// Device/Application/ST/ST_MACHINE/ST_MACHINE_PUBLIC
TYPE ST_MACHINE_PUBLIC :
STRUCT
	xEnabled             : BOOL; // Станок включен в работу
	xDisablePending      : BOOL; // Запрошено отключение после выхода автомата в разрешённый шаг
	xPowerAllowed        : BOOL; // Кнопка включения, отключения или отмены отключения доступна
	xResetAllowed        : BOOL; // Кнопка сброса ошибки станка доступна
	xManualControlAllowed       : BOOL; // Ручное управление разрешено режимом и состоянием станка
	xManualSafetyDoorControlEnabled : BOOL; // Операторская дверь управляется только моделью
	xManualSafetyDoorOpenAllowed : BOOL; // Разрешено открыть операторскую дверь
	xManualSafetyDoorCloseAllowed: BOOL; // Разрешено закрыть операторскую дверь
	xManualHatchOpenAllowed      : BOOL; // Разрешено открыть роботный люк
	xManualHatchCloseAllowed     : BOOL; // Разрешено закрыть роботный люк
	xManualHatchUnlockAllowed    : BOOL; // Разрешено открыть замок роботного люка
	xManualHatchLockAllowed      : BOOL; // Разрешено закрыть замок роботного люка
	xManualChuckOpenAllowed      : BOOL; // Разрешено разжать патрон
	xManualChuckCloseAllowed     : BOOL; // Разрешено зажать патрон
	xProcessing          : BOOL; // Станок выполняет цикл обработки
    xPartReady           : BOOL; // Обработка детали завершена
    xServiceRequired     : BOOL; // Станку требуется обслуживание роботом
    xCanAcceptService    : BOOL; // Станок готов принять робота
    xRobotReleased       : BOOL; // Робот освобождён после операции
	xDone                : BOOL; // Операция обслуживания завершена
    xBusy                : BOOL; // Блок выполняет операцию обслуживания
    xError               : BOOL; // Станок находится в ошибке
	xCriticalError       : BOOL; // Ошибка требует зависимой аварии и остановки робота
	xAlarmError          : BOOL; // Активна первичная ошибка оборудования станка
	xExternalError       : BOOL; // Активна внешняя ошибка
	xServiceRejected     : BOOL; // Обслуживание безопасно отклонено до входа робота в станок
    xDoorOpen            : BOOL; // Дверь станка открыта
    xAlarm               : BOOL; // Активна авария станка
	stIo    			 : ST_MACHINE_IO_STATUS; // Статусы исполнительных механизмов станка
    eRecommendedOperation: E_MACHINE_OPERATION; // Рекомендуемая операция обслуживания
    ePartState           : E_PART_STATE; // Состояние детали в патроне
    ePartType            : E_PART_TYPE; // Тип изделия в патроне: заготовка или готовая деталь
    eAbovePoint          : E_POINT_NAME; // Имя точки над станком
    lrAboveX             : LREAL; // Координата X точки над станком
	tCycleExpected       : TIME; // Ожидаемое время текущего цикла
	tCycleElapsed        : TIME; // Прошедшее время текущего цикла
	tMeasuredCycle       : TIME; // Последнее измеренное время корректного автоцикла
	tRemaining           : TIME; // Оставшееся время обработки
	xCycleTimeValid      : BOOL; // Доступна оценка времени цикла
	xMeasuredTimeValid   : BOOL; // Получено измерение корректного автоцикла
	xCycleOvertime       : BOOL; // Фактический цикл превысил ожидаемое время
END_STRUCT
END_TYPE

// Device/Application/ST/ST_CELL/E_CELL_STATE
{attribute 'qualified_only'}
{attribute 'strict'}
TYPE E_CELL_STATE :
(
	IDLE,
	ROUTE_PAYLOAD,
	SELECT_MACHINE,
	MOVE_TO_MACHINE,
	RELEASE_ROBOT_COMMAND,
	WAIT_MACHINE,
	SERVICE_MACHINE,
	MAGAZINE,
	RELEASE_MAGAZINE,
	WAIT_MAGAZINE,
	ERROR,
	GEOMETRY_WAIT,
	GEOMETRY_TRANSFER
);
END_TYPE

// Device/Application/ST/ST_AXIS_GROUP/ST_AXIS_GROUP_DIAGNOSTICS
TYPE ST_AXIS_GROUP_DIAGNOSTICS :
STRUCT
	iStep            : E_AXIS_GROUP_STATE; // Текущий шаг автомата группы
	iOldStep         : E_AXIS_GROUP_STATE; // Предыдущий шаг автомата
	iNewStep         : E_AXIS_GROUP_STATE; // Новый шаг после перехода
	iPowerMode       : E_AXIS_GROUP_POWER_MODE; // Текущий режим питания группы
    iLastErrorStep   : INT; // Шаг возникновения последней ошибки
    sStepName        : STRING[80]; // Текстовое имя текущего шага
    sWaitReason      : STRING[120]; // Причина ожидания на текущем шаге
    sErrorText       : STRING[120]; // Текст активной ошибки
    sWarningText     : STRING[120]; // Текст активного предупреждения
    stWarning        : ST_WARNING_EVENT; // Последнее предупреждение группы для общего журнала
    tStepPreset      : TIME; // Допустимое время текущего шага
    xStepTimeout     : BOOL; // Превышено допустимое время шага
	xStepChanged     : BOOL; // Шаг изменился в текущем цикле
    udiActualErrorID : UDINT; // Код активной ошибки
    udiLastErrorID   : UDINT; // Код последней ошибки
END_STRUCT
END_TYPE

// Device/Application/ST/ST_POINT_MANAGER/ST_POINT_MANAGER_STATUS
TYPE ST_POINT_MANAGER_STATUS :
STRUCT
	xBusy    : BOOL; // Выполняется проверка точки
	xDone    : BOOL; // Проверка точки завершена
	xInvalid : BOOL; // Точка содержит недопустимые параметры
END_STRUCT
END_TYPE

// Device/Application/GVL/GVL_MAGAZINE
{attribute 'qualified_only'}
VAR_GLOBAL
	astPartStatus : ARRAY [1..2] OF ST_MAGAZINE_STATUS; // Статус только операций робота, без механического обмена
	astAutoCommand : ARRAY [1..GVL_CELL_SETTINGS.MagazineCount] OF ST_MAGAZINE_COMMAND;
	astCommand : ARRAY [1..GVL_CELL_SETTINGS.MagazineCount] OF ST_ROBOT_COMMAND;
	astStatus : ARRAY [1..GVL_CELL_SETTINGS.MagazineCount] OF ST_MAGAZINE_STATUS;
	astDiag : ARRAY [1..GVL_CELL_SETTINGS.MagazineCount] OF ST_MAGAZINE_DIAG;
	astError : ARRAY [1..GVL_CELL_SETTINGS.MagazineCount] OF ST_MAGAZINE_ERRORS;
END_VAR

// Device/Application/GVL/GVL_ROBOT
{attribute 'qualified_only'}
VAR_GLOBAL
	Command       : ST_ROBOT_COMMAND; // Выбранная команда робота
	ModbusCommand : ST_ROBOT_COMMAND; // Команда внешнему роботу
	Status        : ST_ROBOT_STATUS; // Рабочие статусы робота
	Diag          : ST_ROBOT_DIAG; // Состояние автомата робота
	Error         : ST_ROBOT_ERRORS; // Активные и последние ошибки робота
	GripperDiag   : ST_GRIPPER_DIAG; // Диагностика внутреннего блока захвата
	GripperError  : ST_GRIPPER_ERRORS; // Активные и последние ошибки захвата

	xModbusBusy  : BOOL; // Внешний робот выполняет команду
	xModbusDone  : BOOL; // Внешний робот завершил команду
	xModbusError : BOOL; // Ошибка внешнего робота или обмена
END_VAR

// Device/Application/GVL/GVL_MAGAZINE_AXIS
{attribute 'qualified_only'}
VAR_GLOBAL
	// Legacy-объявление оставлено до удаления SoftMotion-узлов Magazine_1/2 через
	// CODESYS. Активная программа массив не читает, не пишет и FB_AXIS для него не создаёт.
	astAxis : ARRAY [1..GVL_CELL_SETTINGS.MagazineCount] OF ST_AXIS;
END_VAR

// Device/Application/GVL/GVL_MACHINE
{attribute 'qualified_only'}
VAR_GLOBAL
	astPhysicalInput : ARRAY [1..3] OF ST_MACHINE_IO_STATUS; // Только ReadPhysicalInputs пишет физическую обратную связь
	Command    : ARRAY [1..3] OF ST_MACHINE_COMMAND; // Команды станков и робота
	Status     : ARRAY [1..3] OF ST_MACHINE_PUBLIC; // Рабочие статусы станков
	Diag       : ARRAY [1..3] OF ST_MACHINE_DIAG; // Состояния автоматов станков
	Error      : ARRAY [1..3] OF ST_MACHINE_ERRORS; // Ошибки станков
END_VAR

// Device/Application/GVL/GVL_POINT_MANAGER
{attribute 'qualified_only'}
VAR_GLOBAL
	PointManager : ST_POINT_MANAGER; // Команды, статусы и диагностика проверки точки
END_VAR

// Device/Application/GVL/GVL_HMI
{attribute 'qualified_only'}
VAR_GLOBAL
	stGeometryRequest : ST_GEOMETRY_REQUEST;
	udiGeometryCommandSeq : UDINT;
	udiGeometryIssuedAtMs : UDINT;
	audiGeometryStopSeq : ARRAY [1..2] OF UDINT;
	{attribute 'symbol' := 'read'}
	audiGeometryStopAck : ARRAY [1..2] OF UDINT;
	{attribute 'symbol' := 'read'}
	udiGeometryAckSeq : UDINT;
	{attribute 'symbol' := 'read'}
	uiGeometryResult : UINT;
	{attribute 'symbol' := 'read'}
	stGeometryCapture : ST_GEOMETRY_CONFIG;
	{attribute 'symbol' := 'read'}
	astGeometryStatus : ARRAY [1..2] OF ST_GEOMETRY_STATUS;
	audiGeometryProducedNormal : ARRAY [1..2] OF UDINT;
	audiGeometryProducedSimulation : ARRAY [1..2] OF UDINT;
	{attribute 'symbol' := 'read'}
	astGeometryConfig : ARRAY [1..2] OF ST_GEOMETRY_CONFIG;
	{attribute 'symbol' := 'read'}
	astGeometryCalls : ARRAY [1..3] OF ST_GEOMETRY_CALL;
	{attribute 'symbol' := 'read'}
	astGeometryEvents : ARRAY [1..100] OF ST_GEOMETRY_EVENT;
	{attribute 'symbol' := 'read'}
	udiGeometryEventSequence : UDINT;
	{attribute 'symbol' := 'read'}
	auiGeometryPeriod : ARRAY [1..3] OF UINT;
	{attribute 'symbol' := 'read'}
	auiGeometryCount : ARRAY [1..3] OF UINT;
	{attribute 'symbol' := 'read'}
	axGeometryCallAllowed : ARRAY [1..3] OF BOOL;
	{attribute 'symbol' := 'read'}
	axGeometryCancelAllowed : ARRAY [1..3] OF BOOL;
	{attribute 'symbol' := 'read'}
	xGeometryAutoEnabled : BOOL;
	{attribute 'symbol' := 'read'}
	xGeometryAutoChangeAllowed : BOOL;
	{attribute 'symbol' := 'read'}
	xGeometrySupported : BOOL;
	{attribute 'symbol' := 'read'}
	xGeometryWaitWhenOccupied : BOOL;
	{attribute 'symbol' := 'read'}
	xGeometrySettingsAllowed : BOOL;
	{attribute 'symbol' := 'read'}
	tGeometryTransportTimeout : TIME;
	{attribute 'symbol' := 'read'}
	tGeometryFeedbackTimeout : TIME;
	{attribute 'symbol' := 'read'}
	tGeometryResetPulse : TIME;
	{attribute 'symbol' := 'read'}
	tGeometryWaitWarningTimeout : TIME;
	{attribute 'symbol' := 'readwrite'}
	stTwinRequest : ST_TWO_PALLET_REQUEST;
	{attribute 'symbol' := 'readwrite'}
	udiTwinCommandSeq : UDINT;
	{attribute 'symbol' := 'readwrite'}
	udiTwinIssuedAtMs : UDINT;
	{attribute 'symbol' := 'read'}
	udiTwinAckSeq : UDINT;
	{attribute 'symbol' := 'read'}
	uiTwinResult : UINT;
	{attribute 'symbol' := 'read'}
	uiMagazineMode : UINT;
	{attribute 'symbol' := 'read'}
	xMagazineModeAllowed : BOOL;
	{attribute 'symbol' := 'read'}
	astTwinStatus : ARRAY [1..2] OF ST_TWO_PALLET_STATUS;
	{attribute 'symbol' := 'read'}
	astTwinConfig : ARRAY [1..2] OF ST_TWO_PALLET_CONFIG;
	{attribute 'symbol' := 'read'}
	astTwinStore : ARRAY [1..2] OF ST_TWO_PALLET_STORE;
	{attribute 'symbol' := 'read'}
	udiHmiCommandClockMs : UDINT;
	{attribute 'symbol' := 'readwrite'}
	audiHmiCommandIssuedAtMs : ARRAY [1..121] OF UDINT;
	{attribute 'symbol' := 'read'}
	auiHmiCommandResult : ARRAY [1..121] OF UINT; // 1 consumed, 2 expired
	{attribute 'symbol' := 'readwrite'}
	udiCellSettingIssuedAtMs : UDINT;
	{attribute 'symbol' := 'readwrite'}
	audiHmiCommandSeq : ARRAY [1..121] OF UDINT;
	{attribute 'symbol' := 'read'}
	audiHmiCommandAckSeq : ARRAY [1..121] OF UDINT;
	{attribute 'symbol' := 'readwrite'}
	uiCellSettingIndex : UINT; // 1..36, see command-contract.mjs
	{attribute 'symbol' := 'readwrite'}
	lrCellSettingRequest : LREAL; // TIME values in milliseconds
	{attribute 'symbol' := 'readwrite'}
	udiCellSettingCommandSeq : UDINT;
	{attribute 'symbol' := 'read'}
	udiCellSettingAckSeq : UDINT;
	{attribute 'symbol' := 'read'}
	uiCellSettingResult : UINT; // 1 applied, 2 blocked, 3 invalid, 4 expired
	{attribute 'symbol' := 'readwrite'}
	uiTestEnvironmentRequest : UINT := UINT#0;
	{attribute 'symbol' := 'read'}
	xTestEnvironmentApply : BOOL;
	{attribute 'symbol' := 'readwrite'}
	uiTestSpeedProfileRequest : UINT := UINT#0;
	{attribute 'symbol' := 'read'}
	xTestSpeedProfileApply : BOOL;
	{attribute 'symbol' := 'readwrite'}
	xTestSessionActive : BOOL;
	{attribute 'symbol' := 'readwrite'}
	xTestAbort : BOOL; // Удерживаемая отмена теста: немедленно прекращает тестовую команду
	{attribute 'symbol' := 'readwrite'}
	stTestScenario : ST_TEST_SCENARIO_BUFFER;
	{attribute 'symbol' := 'read'}
	xTestScenarioApply : BOOL;
	uiTestEnvironmentApplied : UINT;
	uiTestSpeedProfileApplied : UINT;
	xTestEnvironmentChangeAllowed : BOOL;
	xTestScenarioApplyAllowed : BOOL;
	xSc500BenchKeyActive : BOOL; // Устаревшее OPC UA поле, всегда FALSE; физический ключ удалён
	xSc500BenchKeyLost : BOOL; // Устаревшее OPC UA поле, всегда FALSE
	uiTestRejectReason : UINT;
	udiTestScenarioAckSeq : UDINT;
	uiTestScenarioResult : UINT;
	stTestObservability : ST_TEST_OBSERVABILITY;
	{attribute 'symbol' := 'readwrite'}
	xSimulationAccelerationEnable : BOOL := FALSE; // Разрешить ускорение тестовой симуляции
	{attribute 'symbol' := 'readwrite'}
	uiSimulationTimeFactor : UINT := 1; // Запрошенный коэффициент симуляции 1..100
	xSimulationAccelerationActive : BOOL; // Динамика XYZ и таймеры применены с одним коэффициентом
	xSimulationAccelerationChangeAllowed : BOOL; // Ползунок разрешён; изменение ставится в очередь
	uiSimulationTimeFactorApplied : UINT := 1; // Фактически применённый коэффициент
	{attribute 'symbol' := 'read'}
	xSimulationAccelerationPending : BOOL; // Новое значение применится перед следующим тестом
	{attribute 'symbol' := 'read'}
	xSimulationAccelerationBusy : BOOL; // Перенастройка Dynamic Limits выполняется
	xSimulationAccelerationError : BOOL;
	{attribute 'symbol' := 'read'}
	udiSimulationAccelerationErrorId : UDINT;
	{attribute 'symbol' := 'read'}
	lrSafetyHomeX : LREAL := 0.0; // Координата X точки HOME_SAFETY
	{attribute 'symbol' := 'read'}
	lrSafetyHomeY : LREAL := 0.0; // Координата Y точки HOME_SAFETY
	{attribute 'symbol' := 'read'}
	lrSafetyHomeZ : LREAL := 0.0; // Координата Z точки HOME_SAFETY
	{attribute 'symbol' := 'read'}
	lrSafetyHomeSpeedFactor : LREAL := 0.2; // Локальный коэффициент скорости точки 0.1..1.0
	{attribute 'symbol' := 'read'}
	lrSafetyHomeToleranceX : LREAL := 5.0; // Допуск безопасной зоны по X, мм
	{attribute 'symbol' := 'read'}
	lrSafetyHomeToleranceY : LREAL := 5.0; // Допуск безопасной зоны по Y, мм
	{attribute 'symbol' := 'read'}
	lrSafetyHomeToleranceZ : LREAL := 5.0; // Допуск безопасной зоны по Z, мм
	{attribute 'symbol' := 'read'}
	rRobotAccelerationPercent : REAL := 100.0; // Разгон относительно предела осей, 1..100 %
	{attribute 'symbol' := 'read'}
	rRobotDecelerationPercent : REAL := 100.0; // Торможение относительно предела осей, 1..100 %
	{attribute 'symbol' := 'read'}
	rRobotJerkPercent : REAL := 100.0; // Jerk относительно предела осей, 1..100 %
	{attribute 'symbol' := 'read'}
	lrRobotHaltDeceleration : LREAL := 1000.0; // Замедление MC_GroupHalt, мм/с2
	{attribute 'symbol' := 'read'}
	lrRobotHaltJerk : LREAL := 10000.0; // Jerk MC_GroupHalt, мм/с3
	{attribute 'symbol' := 'read'}
	stCellMachineTimeouts : ST_MACHINE_TIMEOUTS; // Настраиваемые TIMEOUT технологических ожиданий
	{attribute 'symbol' := 'read'}
	stCellAxisTimeouts : ST_AXIS_TIMEOUTS; // Общий профиль TIMEOUT осей X/Y/Z
	{attribute 'symbol' := 'read'}
	stCellAxisGroupTimeouts : ST_AXIS_GROUP_TIMEOUTS; // TIMEOUT координатной группы XYZ
	{attribute 'symbol' := 'read'}
	tPointCheckStartTimeout : TIME;
	{attribute 'symbol' := 'read'}
	tSimulationDynamicsTimeout : TIME;
	{attribute 'symbol' := 'read'}
	tHmiWatchdogTimeout : TIME;
	{attribute 'symbol' := 'read'}
	tMobileMotionWatchdogTimeout : TIME;
	{attribute 'symbol' := 'read'}
	tPointCheckWatchdogTimeout : TIME;
	{attribute 'symbol' := 'read'}
	tHmiCommandFreshnessTimeout : TIME;
	{attribute 'symbol' := 'read'}
	tAlarmHornDuration : TIME; // Подтверждённая длительность звука
	tInputFilterRise : TIME := T#20MS;
	{attribute 'symbol' := 'read'}
	tInputFilterFall : TIME := T#20MS;
	{attribute 'symbol' := 'read'}
	xIoFilterSettingsChangeAllowed : BOOL;
	{attribute 'symbol' := 'read'}
	xPhysicalIoActive : BOOL;
	{attribute 'symbol' := 'read'}
	xPhysicalIoMappingVerified : BOOL;
	xCellSettingsChangeAllowed : BOOL; // PLC разрешает изменение настроек ячейки
	// Команды и настройки, получаемые от HMI.
	{attribute 'symbol' := 'read'}
	xCellEnable       : BOOL; // Импульс включения оборудования ячейки
	{attribute 'symbol' := 'read'}
	xCellDisable      : BOOL; // Импульс отключения оборудования ячейки
	{attribute 'symbol' := 'read'}
	xCellStart        : BOOL; // Импульс запуска цикла или отмены ожидающей остановки
	{attribute 'symbol' := 'read'}
	xCellStop         : BOOL; // Импульс остановки автоматического цикла
	{attribute 'symbol' := 'read'}
	xCellReset        : BOOL; // Общий сброс ошибок ячейки
	{attribute 'symbol' := 'read'}
	xSafetyRelayReset : BOOL; // Импульс отдельного сброса реле безопасности
	{attribute 'symbol' := 'readwrite'}
	uiCellOperatorChoice : UINT; // Ответ активному предпусковому опросу PLC
	{attribute 'symbol' := 'read'}
	xCellOperatorChoice : BOOL; // Импульс подтверждения ответа предпускового опроса
	{attribute 'symbol' := 'read'}
	xCellOperatorCancel : BOOL; // Импульс отмены предпускового опроса
	{attribute 'symbol' := 'read'}
	xAlarmResetWarnings : BOOL; // Импульс сброса накопленных предупреждений
	{attribute 'symbol' := 'read'}
	xCellManual       : BOOL; // Фактический режим; единственный писатель — PLC
	{attribute 'symbol' := 'readwrite'}
	xCellManualRequest : BOOL; // Требуемый режим; записать до CommandSeq
	{attribute 'symbol' := 'readwrite'}
	udiCellModeCommandSeq : UDINT; // Новая транзакция переключения режима
	{attribute 'symbol' := 'read'}
	udiCellModeAckSeq : UDINT; // Последняя обработанная транзакция
	{attribute 'symbol' := 'read'}
	uiCellModeResult : UINT; // 0 нет результата, 1 применён, 2 цикл работает, 3 общая авария
	lrOffsetX          : LREAL; // Ручное смещение по оси X
	lrOffsetY          : LREAL; // Ручное смещение по оси Y
	lrOffsetZ          : LREAL; // Ручное смещение по оси Z
	xModbusMode        : BOOL; // Read-only: TRUE, когда PLC применил MODBUS_TCP
	{attribute 'symbol' := 'readwrite'}
	uiRobotControlModeRequest : UINT; // 0 SoftMotion, 1 Modbus TCP
	{attribute 'symbol' := 'read'}
	xRobotControlModeApply : BOOL; // Импульс применения выбранного режима
	{attribute 'symbol' := 'readwrite'}
	uiModbusIpOctet1 : UINT; // Подготавливаемые настройки соединения
	{attribute 'symbol' := 'readwrite'}
	uiModbusIpOctet2 : UINT;
	{attribute 'symbol' := 'readwrite'}
	uiModbusIpOctet3 : UINT;
	{attribute 'symbol' := 'readwrite'}
	uiModbusIpOctet4 : UINT;
	{attribute 'symbol' := 'readwrite'}
	uiModbusPort : UINT := UINT#502;
	{attribute 'symbol' := 'readwrite'}
	uiModbusUnitId : UINT := UINT#1;
	{attribute 'symbol' := 'readwrite'}
	udiModbusResponseTimeoutMs : UDINT := UDINT#500;
	{attribute 'symbol' := 'readwrite'}
	udiModbusPollIntervalMs : UDINT := UDINT#50;
	{attribute 'symbol' := 'readwrite'}
	udiModbusHeartbeatTimeoutMs : UDINT := UDINT#2000;
	{attribute 'symbol' := 'readwrite'}
	udiModbusCommandStartTimeoutMs : UDINT := UDINT#30000;
	{attribute 'symbol' := 'readwrite'}
	udiModbusCommandTimeoutMs : UDINT := UDINT#600000;
	{attribute 'symbol' := 'read'}
	xModbusSettingsApply : BOOL; // Импульс атомарного применения настроек
	xRobotModeChangeAllowed : BOOL;
	xModbusSettingsChangeAllowed : BOOL;
	uiRobotModeRejectReason : UINT; // 0 нет запрета, 1 состояние ячейки, 2 приводы, 3 внешний робот, 4 настройки
	uiModbusSettingsRejectReason : UINT;
	stRobotModbusStatus : ST_ROBOT_MODBUS_STATUS;
	auiRobotModbusWriteRegisters : ARRAY [1..9] OF UINT; // Диагностическая копия 1001..1009, read-only для HMI
	auiRobotModbusReadRegisters : ARRAY [1..17] OF UINT; // Диагностическая копия 1101..1117, read-only для HMI
	{attribute 'symbol' := 'read'}
	xRobotDrivesEnable : BOOL; // Импульс включения приводов робота
	{attribute 'symbol' := 'read'}
	xRobotDrivesDisable: BOOL; // Импульс отключения приводов робота
	{attribute 'symbol' := 'read'}
	xRobotStop         : BOOL; // Импульс контролируемой остановки робота
	{attribute 'symbol' := 'read'}
	xRobotReset        : BOOL; // Импульс сброса ошибок робота и приводов
	{attribute 'symbol' := 'readwrite'}
	udiHmiHeartbeat    : UDINT; // Счётчик связи HMI -> PLC, контролируется PLC watchdog
	{attribute 'symbol' := 'readwrite'}
	xMobileMotionActive : BOOL; // Активная аренда движения от мобильного пульта
	{attribute 'symbol' := 'readwrite'}
	udiMobileMotionHeartbeat : UDINT; // Heartbeat активной мобильной аренды
	xMobileMotionLeaseAlive : BOOL; // Диагностика принятой PLC мобильной аренды
	rMobileMotionAppliedSpeedPercent : REAL; // Защёлкнутый PLC лимит мобильной скорости
	{attribute 'symbol' := 'readwrite'}
	xRobotContinuousMode : BOOL := FALSE; // Режим ручного движения: FALSE шаг, TRUE непрерывный Jog
	{attribute 'symbol' := 'readwrite'}
	rRobotManualSpeedPercent : REAL := 0.1; // Общий override скорости JOG, MoveAbsolute и движения к точкам, 0.1..100 %; имя сохранено для OPC UA
	{attribute 'symbol' := 'readwrite'}
	lrRobotManualStep : LREAL := 1.0; // Шаг короткого относительного перемещения, мм
	// Транзакционный редактор 14 фиксированных инженерных точек.
	{attribute 'symbol' := 'readwrite'}
	uiPointEditorIndex : UINT := UINT#1;
	{attribute 'symbol' := 'readwrite'}
	alrPointEditorDraftXYZ : ARRAY [1..3] OF LREAL;
	{attribute 'symbol' := 'readwrite'}
	lrPointEditorDraftSpeedFactor : LREAL;
	{attribute 'symbol' := 'readwrite'}
	lrPointEditorDraftMagazineSafeZ : LREAL; // Смещение Safe Z базовой точки магазина
	{attribute 'symbol' := 'readwrite'}
	lrPointEditorDraftMagazineChangeZ : LREAL; // Смещение Change Z базовой точки магазина
	{attribute 'symbol' := 'readwrite'}
	uiPointEditorCommand : UINT; // 1 CAPTURE, 2 SAVE, 3 CHECK сохранённой точки
	{attribute 'symbol' := 'readwrite'}
	udiPointEditorCommandSeq : UDINT;
	{attribute 'symbol' := 'readwrite'}
	udiPointCheckHeartbeat : UDINT; // Отдельный heartbeat владельца проверки, не заменяет HMI
	{attribute 'symbol' := 'read'}
	xPointCheckStop : BOOL; // Остановка только текущей проверки, потребляется PLC
	{attribute 'symbol' := 'read'}
	rPointCheckSpeedPercent : REAL := 10.0; // Применённая настройка, 0.1..100 %
	{attribute 'symbol' := 'readwrite'}
	astAxisHmiCommand : ARRAY [1..3] OF ST_AXIS_HMI_COMMAND; // Команды выбранной оси от HMI
	{attribute 'symbol' := 'readwrite'}
	uiRobotManualAction : UINT; // Код E_ROBOT_ACTION без записи типизированного enum через OPC UA
	{attribute 'symbol' := 'readwrite'}
	uiRobotManualPoint : UINT; // Код E_POINT_NAME без записи типизированного enum через OPC UA
	{attribute 'symbol' := 'readwrite'}
	uiRobotManualSlot : UINT := UINT#1; // Активный слот для трёх магазинных точек
	{attribute 'symbol' := 'read'}
	xRobotManualExecute : BOOL; // Импульс ручного действия робота/перехода к точке
	xErrorSimulationEnable : BOOL; // Переключатель диагностического режима эмуляции ошибок
	{attribute 'symbol' := 'read'}
	axSimAxisJogConflict : ARRAY [1..3] OF BOOL; // Импульсы безопасного конфликта Jog осей X/Y/Z
	{attribute 'symbol' := 'read'}
	xSimAxisGroupError : BOOL; // Импульс формирования тестовой ошибки SM3 группы XYZ
	{attribute 'symbol' := 'read'}
	xSimRobotWrongAction : BOOL; // Импульс недопустимого действия робота
	{attribute 'symbol' := 'read'}
	xSimCellBothGrippers : BOOL; // Импульс противоречивого заполнения двух захватов
	xSimGripper1Fault  : BOOL; // Имитация неисправности первого захвата
	xSimGripper2Fault  : BOOL; // Имитация неисправности второго захвата
	xSimGripperRotationFault : BOOL; // Имитация неисправности поворота захвата
	xSimGripperGlobalFault   : BOOL; // Имитация общей неисправности захвата
	{attribute 'symbol' := 'read'}
	xSimPointXOutOfLimit     : BOOL; // Импульс точки с координатой X вне границ
	{attribute 'symbol' := 'read'}
	xSimPointYOutOfLimit     : BOOL; // Импульс точки с координатой Y вне границ
	{attribute 'symbol' := 'read'}
	xSimPointZOutOfLimit     : BOOL; // Импульс точки с координатой Z вне границ
	{attribute 'symbol' := 'read'}
	xSimPointInvalidVelocity : BOOL; // Импульс точки с недопустимой скоростью
	{attribute 'symbol' := 'read'}
	xSimMagazineWrongOperation : BOOL; // Импульс недопустимой операции магазина
	{attribute 'symbol' := 'read'}
	xSimMagazineNoBlank        : BOOL; // Импульс ошибки отсутствия заготовки
	{attribute 'symbol' := 'read'}
	xSimMagazineNoFreeSlot     : BOOL; // Импульс ошибки отсутствия свободного слота
	{attribute 'symbol' := 'read'}
	xSimMagazineInvalidSlot    : BOOL; // Импульс недопустимого номера слота
	{attribute 'symbol' := 'read'}
	xSimMagazineSlotContent    : BOOL; // Импульс несоответствия содержимого слота
	{attribute 'symbol' := 'read'}
	xSimMagazineGeometry       : BOOL; // Импульс недопустимой геометрии магазина
	axSimSafetyEmergencyStopStation : ARRAY [1..4] OF BOOL; // Удерживаемые инъекции грибков постов
	axSimSafetyEmergencyStopCabinet : ARRAY [1..2] OF BOOL; // Удерживаемые инъекции грибков шкафов
	xSimSafetyEmergencyStopMpg : BOOL; // Инъекция грибка MPG-пульта
	xSimSafetyPhaseRelayFault : BOOL; // Инъекция отказа контроля фаз
	xSimSafetyPressureRelayFault : BOOL; // Инъекция отказа контроля давления
	xSimSafetyRelayFault : BOOL; // Инъекция невзведённого реле безопасности
	axSimSafetyDoorUnlocked : ARRAY [1..4] OF BOOL; // Инъекция открытого замка двери
	xMagazineEnable    : BOOL; // Импульс включения магазина
	xMagazineDisable   : BOOL; // Импульс отключения магазина
	xMagazineFillBlanks: BOOL; // Заполнить активные слоты магазина заготовками
	xMagazineClear     : BOOL; // Полностью очистить магазин
	{attribute 'symbol' := 'readwrite'}
	xMagazineCycleSlot : BOOL; // Переключить содержимое выбранного слота
	{attribute 'symbol' := 'readwrite'}
	uiMagazineEditSlot : UINT; // Номер слота, изменяемого оператором
	{attribute 'symbol' := 'readwrite'}
	astMagazineCommand : ARRAY [1..GVL_CELL_SETTINGS.MagazineCount] OF ST_MAGAZINE_HMI_COMMAND;
	{attribute 'symbol' := 'readwrite'}
	uiRobotManualMagazine : UINT := UINT#1; // Магазин ручной роботной команды
	{attribute 'symbol' := 'read'}
	axMachineEnable    : ARRAY [1..3] OF BOOL; // Включить станок или отменить ожидающее отключение
	{attribute 'symbol' := 'read'}
	axMachineDisable   : ARRAY [1..3] OF BOOL; // Импульсы отключения отдельных станков
	{attribute 'symbol' := 'read'}
	axMachineReset     : ARRAY [1..3] OF BOOL; // Команды сброса ошибок отдельных станков
	{attribute 'symbol' := 'read'}
	axMachineManualSafetyDoorOpen  : ARRAY [1..3] OF BOOL; // Ручное открытие операторской двери
	{attribute 'symbol' := 'read'}
	axMachineManualSafetyDoorClose : ARRAY [1..3] OF BOOL; // Ручное закрытие операторской двери
	{attribute 'symbol' := 'read'}
	axMachineManualHatchOpen       : ARRAY [1..3] OF BOOL; // Ручное открытие роботного люка
	{attribute 'symbol' := 'read'}
	axMachineManualHatchClose      : ARRAY [1..3] OF BOOL; // Ручное закрытие роботного люка
	{attribute 'symbol' := 'read'}
	axMachineManualHatchUnlock     : ARRAY [1..3] OF BOOL; // Ручное открытие замка роботного люка
	{attribute 'symbol' := 'read'}
	axMachineManualHatchLock       : ARRAY [1..3] OF BOOL; // Ручное закрытие замка роботного люка
	{attribute 'symbol' := 'read'}
	axMachineManualChuckOpen       : ARRAY [1..3] OF BOOL; // Ручной разжим патрона
	{attribute 'symbol' := 'read'}
	axMachineManualChuckClose      : ARRAY [1..3] OF BOOL; // Ручной зажим патрона
	{attribute 'symbol' := 'read'}
	axMachineSimReset  : ARRAY [1..3] OF BOOL; // Отдельный сброс аварий FB_MACHINE_SIMULATION
	axMachineSimAlarm  : ARRAY [1..3] OF BOOL; // Имитация общей аварии станков
	axMachineSimDoorFault  : ARRAY [1..3] OF BOOL; // Имитация неисправности роботных люков
	{attribute 'symbol' := 'readwrite'}
	axMachineSimSafetyDoorOpen : ARRAY [1..3] OF BOOL; // Имитация открытой операторской двери
	axMachineSimChuckFault : ARRAY [1..3] OF BOOL; // Имитация неисправности патронов станков
	axMachineTimeoutRobotMove    : ARRAY [1..3] OF BOOL; // Игнорировать завершение движения робота до TIMEOUT
	axMachineTimeoutRobotAction  : ARRAY [1..3] OF BOOL; // Игнорировать завершение действия захвата до TIMEOUT
	axMachineTimeoutRobotRelease : ARRAY [1..3] OF BOOL; // Игнорировать освобождение интерфейса робота до TIMEOUT
	axMachineTimeoutDoorOpen     : ARRAY [1..3] OF BOOL; // Игнорировать подтверждение открытия двери до TIMEOUT
	axMachineTimeoutDoorClose    : ARRAY [1..3] OF BOOL; // Игнорировать подтверждение закрытия двери до TIMEOUT
	axMachineTimeoutHatchUnlock  : ARRAY [1..3] OF BOOL; // Игнорировать подтверждение открытия замка до TIMEOUT
	axMachineTimeoutChuckOpen    : ARRAY [1..3] OF BOOL; // Игнорировать подтверждение разжима патрона до TIMEOUT
	axMachineTimeoutChuckClose   : ARRAY [1..3] OF BOOL; // Игнорировать подтверждение зажима патрона до TIMEOUT
	axMachineTimeoutCycleStart   : ARRAY [1..3] OF BOOL; // Игнорировать подтверждение запуска цикла до TIMEOUT
	{attribute 'symbol' := 'read'}
	axMachineSetBlank  : ARRAY [1..3] OF BOOL; // Подтвердить заготовку в патроне
	{attribute 'symbol' := 'read'}
	axMachineSetDetail : ARRAY [1..3] OF BOOL; // Подтвердить готовую деталь в патроне
	{attribute 'symbol' := 'read'}
	axMachineAcceptDoor: ARRAY [1..3] OF BOOL; // Подтвердить закрытие двери
	{attribute 'symbol' := 'read'}
	axMachineRejectDoor: ARRAY [1..3] OF BOOL; // Отказаться от закрытия двери
	{attribute 'symbol' := 'read'}
	axMachineAcceptRun : ARRAY [1..3] OF BOOL; // Подтвердить запуск обработки
	{attribute 'symbol' := 'read'}
	axMachineRejectRun : ARRAY [1..3] OF BOOL; // Отказаться от запуска обработки
	axMachineUsed      : ARRAY [1..3] OF BOOL := [FALSE, FALSE, FALSE]; // Выбор станков для авто; FB_MACHINE после старта находится в DISABLED
	xUseHmiCycleTime   : ARRAY [1..3] OF BOOL := [FALSE, FALSE, FALSE]; // Использовать заданное время цикла
	tMachineCycleTime  : ARRAY [1..3] OF TIME := [T#60S, T#60S, T#60S]; // Время цикла станков
	tMachineDoorOpenTime   : TIME := T#1S; // Время открытия люка в симуляторе станка
	tMachineDoorCloseTime  : TIME := T#1S; // Время закрытия люка в симуляторе станка
	tMachineChuckOpenTime  : TIME := T#1S; // Время разжима патрона в симуляторе станка
	tMachineChuckCloseTime : TIME := T#1S; // Время зажима патрона в симуляторе станка
	tGripper1OpenTime   : TIME := T#500MS; // Время открытия первого захвата
	tGripper1CloseTime  : TIME := T#500MS; // Время закрытия первого захвата
	tGripper2OpenTime   : TIME := T#500MS; // Время открытия второго захвата
	tGripper2CloseTime  : TIME := T#500MS; // Время закрытия второго захвата
	tGripperChangeTime  : TIME := T#700MS; // Время смены рабочего захвата
	{attribute 'symbol' := 'read'}
	MagazineRows       : UINT := 12; // Статичная кассета: 12 рядов
	{attribute 'symbol' := 'read'}
	MagazineColumns    : UINT := 10; // Число столбцов магазина
	{attribute 'symbol' := 'read'}
	MagazinePitchX     : LREAL := 60.0; // Шаг слотов по оси X
	{attribute 'symbol' := 'read'}
	MagazinePitchY     : LREAL := 60.0; // Шаг слотов по оси Y
	stRobotCommand     : ST_ROBOT_COMMAND; // Ручная команда роботу или магазину
	{attribute 'symbol' := 'readwrite'}
	stMultiType        : ST_MULTI_TYPE_HMI; // Конфигурация типов и диагностика универсального цикла

	// Данные, передаваемые в HMI.
	udiPlcHeartbeat : UDINT; // Счётчик циклов PLC для контроля связи
	xHmiConnectionAlive : BOOL; // PLC видит актуальный heartbeat HMI
	xManualRecoveryActive : BOOL; // Разрешён ограниченный Jog в режиме восстановления
	astAxisHmiStatus : ARRAY [1..3] OF ST_AXIS_HMI_STATUS; // xAllowed и диагностика ручного управления по осям
	stRobotHmiStatus : ST_ROBOT_HMI_STATUS; // xAllowed и диагностика ручных действий робота
	xGlobalError    : BOOL; // Активна общая ошибка ячейки
	xErrorSimulationEnabled : BOOL; // Фактическое состояние диагностического режима
	xSimAxisGroupErrorAllowed : BOOL; // Разрешена безопасная инъекция ошибки SM3
	astAxisFaultStatus : ARRAY [1..3] OF ST_FAULT_INJECTION_STATUS; // Доступность инъекции осей X/Y/Z
	stAxisGroupFaultStatus : ST_FAULT_INJECTION_STATUS; // Состояние инжектора SM3 группы
	stGripperFaultStatus   : ST_FAULT_INJECTION_STATUS; // Состояние инжектора захвата
	stRobotFaultStatus     : ST_FAULT_INJECTION_STATUS; // Состояние локального инжектора робота
	stCellFaultStatus      : ST_FAULT_INJECTION_STATUS; // Состояние инжектора менеджера ячейки
	stSafetyFaultStatus    : ST_FAULT_INJECTION_STATUS; // Состояние инжектора дискретной безопасности
	stPointFaultStatus     : ST_FAULT_INJECTION_STATUS; // Состояние инжектора проверки точки
	stMagazineFaultStatus  : ST_FAULT_INJECTION_STATUS; // Legacy: первый магазин
	astMagazineFaultStatus : ARRAY [1..GVL_CELL_SETTINGS.MagazineCount] OF ST_FAULT_INJECTION_STATUS;
	astMachineFaultStatus  : ARRAY [1..3] OF ST_FAULT_INJECTION_STATUS; // Источники аварий станков
	astMachineTimeouts     : ARRAY [1..3] OF ST_MACHINE_TIMEOUTS; // Действующие таймауты станков
	lrActualX       : LREAL; // Текущая координата X
	lrActualY       : LREAL; // Текущая координата Y
	lrActualZ       : LREAL; // Текущая координата Z
	astPointEditorPoints : ARRAY [1..14] OF ST_POINT; // Прежние 12 точек и базы ГК 1/2
	auiPointEditorPointId : ARRAY [1..14] OF UINT; // Фактические числовые E_POINT_NAME
	stPointEditorResultPoint : ST_POINT; // Результат Capture либо подтверждённого Save
	udiPointEditorAckSeq : UDINT; // Последняя обработанная транзакция
	uiPointEditorResult : UINT; // 0 ожидание, 1 выполнено, 2 отклонено
	uiPointEditorRejectReason : UINT; // Подробная причина отклонения для HMI
	xPointEditorCaptureAllowed : BOOL; // Авторитетное разрешение PLC на Capture
	xPointEditorSaveAllowed : BOOL; // Авторитетное разрешение PLC на Save
	axPointCheckAllowed : ARRAY [1..14] OF BOOL;
	auiPointCheckRejectReason : ARRAY [1..14] OF UINT;
	xPointCheckActive : BOOL;
	uiPointCheckIndex : UINT;
	uiPointCheckState : UINT; // 0 idle, 1 running, 2 completed, 3 stopped, 4 failed
	udiPointCheckRunSeq : UDINT; // Транзакция, которой принадлежит состояние проверки
	rPointCheckAppliedSpeedPercent : REAL := 10.0;
	xPointTableReady : BOOL; // Все 12 базовых точек настроены
	{attribute 'symbol' := 'read'}
	rLoadCNC_1      : REAL; // Процент загрузки станка 1
	{attribute 'symbol' := 'read'}
	rLoadCNC_2      : REAL; // Процент загрузки станка 2
	{attribute 'symbol' := 'read'}
	rLoadCNC_3      : REAL; // Процент загрузки станка 3
	{attribute 'symbol' := 'read'}
	rRobot          : REAL; // Процент загрузки робота

	stCellStatus : ST_CELL_STATUS; // Рабочее состояние автоматического цикла
	stCellDiag   : ST_CELL_DIAG; // Текущий шаг менеджера ячейки
	stCellError  : ST_CELL_ERRORS; // Активные и последние ошибки менеджера ячейки
	stCellSafetyStatus : ST_CELL_SAFETY_STATUS; // Готовность грибков, реле и дверей
	stCellSafetyDiag   : ST_CELL_SAFETY_DIAG; // Отклонённые команды безопасности
	stCellSafetyError  : ST_CELL_SAFETY_ERRORS; // Отдельные Safety-аварии
	{attribute 'symbol' := 'read'}
	astButtonStationIoStatus : ARRAY [1..4] OF ST_BUTTON_STATION_IO_STATUS;
	stFrontControlCabinetIoStatus : ST_CONTROL_CABINET_IO_STATUS;
	{attribute 'symbol' := 'read'}
	xSignalTowerRed   : BOOL; // Фактический логический выход красной секции, включая мигание
	{attribute 'symbol' := 'read'}
	xSignalTowerAmber : BOOL; // Фактический логический выход оранжевой секции
	{attribute 'symbol' := 'read'}
	xSignalTowerGreen : BOOL; // Фактический логический выход зелёной секции, включая мигание
	stRearControlCabinetIoStatus : ST_CONTROL_CABINET_IO_STATUS;
	stMpgIoStatus : ST_MPG_IO_STATUS;
	astEnclosureDoorStatus : ARRAY [1..4] OF ST_ENCLOSURE_DOOR_STATUS;

	stRobotStatus : ST_ROBOT_STATUS; // Состояние робота и двух захватов
	stRobotDiag   : ST_ROBOT_DIAG; // Текущее действие и целевая точка робота
	stRobotError  : ST_ROBOT_ERRORS; // Активные и последние ошибки робота
	stGripperDiag : ST_GRIPPER_DIAG; // Диагностика внутреннего симулятора захвата
	stGripperError: ST_GRIPPER_ERRORS; // Активные и последние ошибки симулятора захвата
	stAxisGroupStatus : ST_AXIS_GROUP_STATUS; // Статусы группы XYZ, включая разрешение тестовой ошибки
	stAxisGroupDiag   : ST_AXIS_GROUP_DIAGNOSTICS; // Диагностика и ErrorID группы XYZ
	stAxisGroupError  : ST_AXIS_GROUP_ERRORS; // Активные и последние ошибки группы XYZ
	astAxisStatus : ARRAY [1..3] OF ST_AXIS_STATUS; // Статусы осей X/Y/Z
	astAxisDiag   : ARRAY [1..3] OF ST_AXIS_DIAGNOSTICS; // Диагностика осей X/Y/Z
	astAxisError  : ARRAY [1..3] OF ST_AXIS_ERROR_CODES; // Ошибки осей X/Y/Z
	stMotionManagerStatus : ST_MOTION_MANAGER_STATUS; // Состояние менеджера движения
	stMotionManagerDiag   : ST_MOTION_MANAGER_DIAG; // Диагностика менеджера движения
	stMotionManagerError  : ST_MOTION_MANAGER_ERRORS; // Ошибки менеджера движения
	stPointManagerStatus  : ST_POINT_MANAGER_STATUS; // Состояние проверки точки
	stPointManagerDiag    : ST_POINT_MANAGER_DIAG; // Диагностика проверки точки
	stPointManagerError   : ST_POINT_MANAGER_ERRORS; // Ошибки проверки точки

	{attribute 'symbol' := 'read'}
	astMachineStatus   : ARRAY [1..3] OF ST_MACHINE_PUBLIC; // Рабочие состояния станков
	astMachineIoStatus : ARRAY [1..3] OF ST_MACHINE_IO_STATUS; // Двери, замки, патроны и циклы станков
	astMachineRawIoStatus : ARRAY [1..3] OF ST_MACHINE_IO_STATUS; // Обратная связь до инжектора
	astMachineDiag     : ARRAY [1..3] OF ST_MACHINE_DIAG; // Текущие шаги и операции станков
	astMachineError    : ARRAY [1..3] OF ST_MACHINE_ERRORS; // Активные и последние ошибки станков
	astMachineSimDiag  : ARRAY [1..3] OF ST_MACHINE_SIM_DIAG; // Диагностика симуляторов станков
	astMachineSimError : ARRAY [1..3] OF ST_MACHINE_SIM_ERRORS; // Ошибки симуляторов станков

	{attribute 'symbol' := 'read'}
	stMagazineStatus : ST_MAGAZINE_STATUS; // Legacy: первый магазин
	stMagazineDiag   : ST_MAGAZINE_DIAG;
	stMagazineError  : ST_MAGAZINE_ERRORS;
	astMagazineSlot  : ARRAY [1..GVL_CELL_SETTINGS.NumberDetail] OF ST_DETAIL;
	astMagazineStatus : ARRAY [1..GVL_CELL_SETTINGS.MagazineCount] OF ST_MAGAZINE_STATUS;
	astMagazineDiag : ARRAY [1..GVL_CELL_SETTINGS.MagazineCount] OF ST_MAGAZINE_DIAG;
	astMagazineError : ARRAY [1..GVL_CELL_SETTINGS.MagazineCount] OF ST_MAGAZINE_ERRORS;
	astMagazineInventory : ARRAY [1..GVL_CELL_SETTINGS.MagazineCount] OF ST_MAGAZINE_INVENTORY;
	stAlarmStatus : ST_ALARM_STATUS; // Сводный статус аварий и предупреждений
	astAlarmEvent : ARRAY [1..100] OF ST_ALARM_EVENT; // Журнал активных и зафиксированных событий


    {attribute 'symbol' := 'read'}
    xIoDoOverrideAllowed : BOOL;
    {attribute 'symbol' := 'read'}
    xIoManualControlActive : BOOL;
    {attribute 'symbol' := 'read'}
    xIoManualStartAllowed : BOOL;
    {attribute 'symbol' := 'read'}
    uiIoDoBlockReason : UINT;
    {attribute 'symbol' := 'read'}
    adwIoDoAllowed : ARRAY [1..2] OF DWORD;
    {attribute 'symbol' := 'read'}
    adwIoDoOnAllowed : ARRAY [1..2] OF DWORD;
    {attribute 'symbol' := 'read'}
    adwIoForcedDo : ARRAY [1..2] OF DWORD;
    {attribute 'symbol' := 'read'}
    adwIoInhibitedDo : ARRAY [1..2] OF DWORD;
    {attribute 'symbol' := 'read'}
    xIoEmergencyStopActive : BOOL;
    {attribute 'symbol' := 'read'}
    xIoEmergencyResetAllowed : BOOL;
    {attribute 'symbol' := 'readwrite'}
    uiIoEmergencyAction : UINT; // 1 остановить; 2 снять программный останов
    {attribute 'symbol' := 'readwrite'}
    udiIoEmergencyIssuedAtMs : UDINT;
    {attribute 'symbol' := 'readwrite'}
    udiIoEmergencyCommandSeq : UDINT;
    {attribute 'symbol' := 'read'}
    udiIoEmergencyAckSeq : UDINT;
    {attribute 'symbol' := 'read'}
    uiIoEmergencyResult : UINT;

    // Физическая диагностика. Команда — payload, время, затем Seq; статусы только чтение.
    {attribute 'symbol' := 'readwrite'}
    uiIoOverrideIndex : UINT;
    {attribute 'symbol' := 'readwrite'}
    uiIoOverrideAction : UINT; // 1..3 DI; 4..6 DO; 7 вернуть всё программе; 8 включить ручное I/O; 9 завершить ручное I/O
    {attribute 'symbol' := 'readwrite'}
    xIoOverrideValue : BOOL;
    {attribute 'symbol' := 'readwrite'}
    udiIoOverrideIssuedAtMs : UDINT;
    {attribute 'symbol' := 'readwrite'}
    udiIoOverrideCommandSeq : UDINT;
    {attribute 'symbol' := 'readwrite'}
    udiIoOverrideHeartbeat : UDINT; // Только открытая страница I/O; watchdog 3 с
    {attribute 'symbol' := 'readwrite'}
    udiIoOverrideHeartbeatAtMs : UDINT; // Время PLC, при STOP не превращает старый heartbeat в новую аренду
    {attribute 'symbol' := 'read'}
    udiIoOverrideAckSeq : UDINT;
    {attribute 'symbol' := 'read'}
    uiIoOverrideResult : UINT; // 1 применено; 2 запрещено; 3 некорректно; 4 просрочено
    {attribute 'symbol' := 'read'}
    xIoOverrideAllowed : BOOL;
    {attribute 'symbol' := 'read'}
    uiIoOverrideBlockReason : UINT; // 0 ручное I/O активно; 2 не ручной режим; 3 нет останова для входа; 7 включите ручное I/O
    {attribute 'symbol' := 'read'}
    uiIoForcedCount : UINT;
    {attribute 'symbol' := 'read'}
    adwIoRawDi : ARRAY [1..3] OF DWORD;
    {attribute 'symbol' := 'read'}
    adwIoUsedDi : ARRAY [1..3] OF DWORD;
    {attribute 'symbol' := 'read'}
    adwIoForcedDi : ARRAY [1..3] OF DWORD;
    {attribute 'symbol' := 'read'}
    adwIoDo : ARRAY [1..2] OF DWORD;
    {attribute 'symbol' := 'read'}
    asIoJournal : ARRAY [1..100] OF STRING(96); // Seq;мс;DI/DO;index;kind;old;new
    {attribute 'symbol' := 'read'}
    udiIoJournalRevision : UDINT; // Seqlock: нечётный — запись, чётный — целостный FIFO
    {attribute 'symbol' := 'read'}
    udiIoJournalSequence : UDINT;
    {attribute 'symbol' := 'read'}
    uiIoJournalHead : UINT;
    {attribute 'symbol' := 'read'}
    uiIoJournalCount : UINT;
    {attribute 'symbol' := 'read'}
    sIoClockMs : STRING(24);

	// Совместимость с существующей визуализацией до штатного обновления XML.
	HMI : ST_HMI; // Старый путь GVL_HMI.HMI.ActualX/Y/Z
END_VAR

VAR_GLOBAL RETAIN
    {attribute 'symbol' := 'read'}
    udiIoBootCounter : UDINT; // Меняется при старте приложения; подмены и FIFO не RETAIN
END_VAR

// Device/Application/GVL/GVL_AXIS_GROUP
{attribute 'qualified_only'}
VAR_GLOBAL
	AxisGroup : ST_AXIS_GROUP; // Команды, статусы и диагностика группы XYZ
END_VAR

// Device/Application/GVL/GVL_ROBOT_MODBUS
{attribute 'qualified_only'}
VAR_GLOBAL
	xModeActive             : BOOL; // TRUE, когда применён MODBUS_TCP
	xRobotModeChangeAllowed : BOOL; // Авторитетное разрешение PLC
	xSettingsChangeAllowed  : BOOL; // Авторитетное разрешение PLC
	xReconnectRequest       : BOOL; // Одноцикловый запрос переподключения клиента
	Config                  : ST_ROBOT_MODBUS_CONFIG;
	Status                  : ST_ROBOT_MODBUS_STATUS;
	Command                 : ST_ROBOT_COMMAND;
	auiWriteRegisters       : ARRAY [0..8] OF UINT; // 1001..1009
	auiReadRegisters        : ARRAY [0..16] OF UINT; // 1101..1117
END_VAR

// Device/Application/GVL/GVL_CELL_CONTROL
{attribute 'qualified_only'}
VAR_GLOBAL
	xGlobalError : BOOL; // Глобальная ошибка ячейки
	xReset       : BOOL; // Общий сброс ошибок ячейки
	xManual      : BOOL; // Ручной режим управления ячейкой
	xEnable      : BOOL; // Импульс включения оборудования ячейки
	xDisable     : BOOL; // Импульс отключения оборудования ячейки
	xStart       : BOOL; // Импульс запуска цикла или отмены ожидающей остановки
	xStop        : BOOL; // Импульс остановки автоматического цикла
END_VAR

// Device/Application/GVL/GVL_CELL_MANAGER
{attribute 'qualified_only'}
VAR_GLOBAL
	Command : ST_CELL_COMMAND; // Команды менеджера ячейки
	Status  : ST_CELL_STATUS; // Рабочие статусы ячейки
	Diag    : ST_CELL_DIAG; // Состояние автомата ячейки
	Error   : ST_CELL_ERRORS; // Ошибки менеджера ячейки
END_VAR

// Device/Application/GVL/GVL_POINT
{attribute 'qualified_only'}
VAR_GLOBAL
	Points : ARRAY [0..iPointNumber] OF ST_POINT; // Глобальная таблица именованных точек
END_VAR

VAR_GLOBAL PERSISTENT RETAIN
	// Постоянное хранилище базовых точек в энергонезависимой памяти контроллера.
	// Размер 15 сохранён ради совместимости со старой раскладкой: позиции 2, 6 и 10
	// (legacy MACHINE_x_INSIDE) больше не публикуются и не участвуют в готовности.
	astRetainPoints : ARRAY [1..iPersistentPointCapacity] OF ST_POINT;
	udiPointStorageVersion : UDINT;
END_VAR

VAR_GLOBAL CONSTANT 
	iPointNumber : INT := 100; // Максимальный индекс таблицы точек
	iEditablePointCount : INT := 14; // 12 прежних точек и 2 базы ГК
	iRequiredPointCount : INT := 12; // ГК проверяет свою настройку при включении станции
	iPersistentPointCapacity : INT := 15;
	udiExpectedPointStorageVersion : UDINT := UDINT#1;
END_VAR

// Device/Application/GVL/GVL_ALARM
{attribute 'qualified_only'}
VAR_GLOBAL
	Command : ST_ALARM_COMMAND; // Команды управления журналом аварий
	Status  : ST_ALARM_STATUS; // Сводный статус аварий и предупреждений
	Events  : ARRAY [1..100] OF ST_ALARM_EVENT; // Кольцевой журнал событий
END_VAR

// Device/Application/GVL/GVL_STATISTIC
{attribute 'qualified_only'}
VAR_GLOBAL
	stStatistic			: ST_STATISTIC;
END_VAR

// Device/Application/GVL/GVL_ROBOT_MODBUS_RETAIN
{attribute 'qualified_only'}
VAR_GLOBAL RETAIN
	eControlMode      : E_ROBOT_CONTROL_MODE := E_ROBOT_CONTROL_MODE.SOFTMOTION;
	aIpAddress        : ARRAY [0..3] OF BYTE := [BYTE#0, BYTE#0, BYTE#0, BYTE#0];
	uiPort            : UINT := UINT#502;
	uiUnitId          : UINT := UINT#1;
	tResponseTimeout  : TIME := T#500MS;
	tPollInterval     : TIME := T#50MS;
	tHeartbeatTimeout : TIME := T#2S;
	tCommandStartTimeout : TIME := T#30S;
	tCommandTimeout   : TIME := T#600S;
END_VAR

// Device/Application/GVL/GVL_CELL_SAFETY_IO
{attribute 'qualified_only'}
VAR_GLOBAL
	// Логические точки для назначения в Device I/O Mapping. Полярность НЗ-контактов
	// нормализуется при привязке: здесь TRUE всегда означает указанное состояние.
	// Начальное состояние стенда: двери закрыты, грибки отжаты, реле в норме.
	axDoorLockClosedInput : ARRAY [1..4] OF BOOL := [TRUE, TRUE, TRUE, TRUE];
	axDoorUnlockButtonInput : ARRAY [1..4] OF BOOL := [FALSE, FALSE, FALSE, FALSE];
	axEmergencyStopButtonStationInput : ARRAY [1..4] OF BOOL := [FALSE, FALSE, FALSE, FALSE];
	// Виртуальные входы постов: учитываются только в среде SIMULATION.
	axSimDoorUnlockButtonInput : ARRAY [1..4] OF BOOL := [FALSE, FALSE, FALSE, FALSE];
	axSimEmergencyStopButtonStationInput : ARRAY [1..4] OF BOOL := [FALSE, FALSE, FALSE, FALSE];
	axEmergencyStopCabinetInput : ARRAY [1..2] OF BOOL := [FALSE, FALSE];
	xEmergencyStopMpgInput : BOOL := FALSE;
	xPhaseRelayOkInput    : BOOL := TRUE;
	xPressureRelayOkInput : BOOL := TRUE;
	xSafetyRelayOkInput   : BOOL := TRUE;
	xCellStartButtonInput : BOOL := FALSE;
	xCellStopButtonInput  : BOOL := FALSE;
	xCellResetButtonInput : BOOL := FALSE;
	xMpgAxisXInput : BOOL := FALSE;
	xMpgAxisYInput : BOOL := FALSE;
	xMpgAxisZInput : BOOL := FALSE;
	xMpgMultiplier1Input : BOOL := FALSE;
	xMpgMultiplier10Input : BOOL := FALSE;
	xMpgMultiplier100Input : BOOL := FALSE;

	// Выходы для назначения на физические каналы.
	axDoorUnlockOutput : ARRAY [1..4] OF BOOL;
	axDoorButtonLampOutput : ARRAY [1..4] OF BOOL;
	xSafetyRelayResetOutput : BOOL;
	// Светосигнальная колонна: готовые уровни с миганием из PLC_PRG.RunSignalTower.
	xAlarmHornOutput : BOOL; // Короткий звук при новой аварии
	xSignalTowerRedOutput   : BOOL;
	xSignalTowerAmberOutput : BOOL;
	xSignalTowerGreenOutput : BOOL;
END_VAR

// Device/Application/GVL/GVL_GEOMETRY_CONTROL
{attribute 'qualified_only'}
VAR_GLOBAL
	astStatus : ARRAY [1..2] OF ST_GEOMETRY_STATUS;
	astSignals : ARRAY [1..2] OF ST_GEOMETRY_SIGNALS;
	astActiveConfig : ARRAY [1..2] OF ST_GEOMETRY_CONFIG;
	astActiveMemory : ARRAY [1..2] OF ST_GEOMETRY_MEMORY;
	astCalls : ARRAY [1..3] OF ST_GEOMETRY_CALL;
	astSimulationConfig : ARRAY [1..2] OF ST_GEOMETRY_CONFIG;
	astSimulationMemory : ARRAY [1..2] OF ST_GEOMETRY_MEMORY;
	astSimulationCalls : ARRAY [1..3] OF ST_GEOMETRY_CALL;
	axSimulationAlarm : ARRAY [1..2] OF BOOL;
	auiAction : ARRAY [1..2] OF UINT;
	astWarning : ARRAY [1..2] OF ST_WARNING_EVENT;
	stCellWarning : ST_WARNING_EVENT;
	astEvents : ARRAY [1..100] OF ST_GEOMETRY_EVENT;
	uiLastStation : UINT;
	uiEnvironment : UINT;
	xSupported : BOOL;
	xAutoChangeAllowed : BOOL;
	xSettingsAllowed : BOOL;
	axCallAllowed : ARRAY [1..3] OF BOOL;
	axCancelAllowed : ARRAY [1..3] OF BOOL;
	auiActiveCount : ARRAY [1..3] OF UINT;
	auiSimulationCount : ARRAY [1..3] OF UINT;
END_VAR
VAR_GLOBAL PERSISTENT RETAIN
	astConfig : ARRAY [1..2] OF ST_GEOMETRY_CONFIG;
	astMemory : ARRAY [1..2] OF ST_GEOMETRY_MEMORY;
	astRetainCalls : ARRAY [1..3] OF ST_GEOMETRY_CALL;
	udiNextCallId : UDINT;
	udiEventSequence : UDINT;
	xAutoEnabled : BOOL := FALSE;
	auiPeriod : ARRAY [1..3] OF UINT := [20, 20, 20];
	auiCount : ARRAY [1..3] OF UINT;
	xWaitWhenOccupied : BOOL := TRUE;
	tTransportTimeout : TIME := T#10S;
	tDriveFeedbackTimeout : TIME := T#3S;
	tResetPulse : TIME := T#1S;
	tWaitWarningTimeout : TIME := T#180S; // Ожидание готовой вызванной детали в станке до WARNING
END_VAR

// Device/Application/GVL/GVL_TEST_IO
{attribute 'qualified_only'}
VAR_GLOBAL
	// Физический ключ стенда исключён из схемы. GVL оставлена для совместимости дерева проекта.
END_VAR

// Device/Application/GVL/GVL_CELL_SETTINGS
{attribute 'qualified_only'}
VAR_GLOBAL CONSTANT
	MagazineCount : INT := 2; // Два независимых статичных магазина
	MagazineSlots : SINT := 120; // Одна кассета 12 x 10 в каждом магазине
	NumberDetail : SINT := 120;
END_VAR

VAR_GLOBAL
	MagazineRows : UINT := 12;
	MagazineColumns : UINT := 10;
	// Не RETAIN: после каждого запуска PLC тестовая среда всегда SIMULATION.
	eTestEnvironment : E_CELL_TEST_ENVIRONMENT := E_CELL_TEST_ENVIRONMENT.SIMULATION;
	eTestSpeedProfile : E_TEST_SPEED_PROFILE := E_TEST_SPEED_PROFILE.REALTIME;
	xSimulationAccelerationEnable : BOOL := FALSE; // Ускорять таймеры и динамику SoftMotion в тестовом профиле FAST
	uiSimulationTimeFactor : UINT := 1; // Запрошенный коэффициент 1..100; можно менять в любой момент
	xSimulationAccelerationActive : BOOL := FALSE; // Применён ускоренный комплект лимитов и таймеров
	uiSimulationTimeFactorApplied : UINT := 1; // Коэффициент, подтверждённый транзакцией Dynamic Limits
	xSimulationAccelerationChangeAllowed : BOOL := FALSE; // Разрешено запомнить новое требование из HMI
	xSimulationAccelerationPending : BOOL := FALSE; // Новое значение ждёт следующего теста
	xSimulationAccelerationBusy : BOOL := FALSE; // Stop/Disable/Change/Enable выполняется
	xSimulationAccelerationError : BOOL := FALSE;
	udiSimulationAccelerationErrorId : UDINT := UDINT#0;
	xErrorSimulationEnabled : BOOL := FALSE; // Разрешение диагностической инъекции ошибок из HMI

	// Безопасный повторный запуск после аварийной остановки.
	// Погрешности задают допустимый диапазон относительно точки HOME_SAFETY.
	lrSafetyHomeToleranceX : LREAL := 5.0;
	lrSafetyHomeToleranceY : LREAL := 5.0;
	lrSafetyHomeToleranceZ : LREAL := 5.0;
	rPointCheckSpeedPercent : REAL := 10.0; // Скорость проверки точки с телефона
	// Допуск контроля неизменности позы после штатной остановки защищает от
	// дрожания обратной связи, но фиксирует последующее ручное перемещение.
	lrStoppedPoseTolerance : LREAL := 1.0;

	// Общий профиль динамики SoftMotion. Проценты масштабируют фактические
	// динамические пределы каждой оси; Halt-параметры принадлежат группе XYZ.
	rRobotAccelerationPercent : REAL := 100.0;
	rRobotDecelerationPercent : REAL := 100.0;
	rRobotJerkPercent : REAL := 100.0;
	lrRobotHaltDeceleration : LREAL := 1000.0;
	lrRobotHaltJerk : LREAL := 10000.0;

	// Настройки ячейки редактируются из HMI только в остановленном безопасном состоянии.
	xCellSettingsChangeAllowed : BOOL := FALSE;
	xIoFilterSettingsChangeAllowed : BOOL := FALSE; // Разрешение фильтров и длительности гудка; применимо и в Modbus
	tAlarmHornDuration : TIME := T#2S; // Звук новой аварии 0..60 с; 0 отключает звук
	tInputFilterRise : TIME := T#20MS; // Стабильный передний фронт обычных DI, 0..5000 мс
	tInputFilterFall : TIME := T#20MS; // Стабильный задний фронт обычных DI, 0..5000 мс
	stMachineTimeouts : ST_MACHINE_TIMEOUTS := (
		tRobotMove := T#60S,
		tRobotAction := T#10S,
		tRobotRelease := T#5S,
		tDoorOpen := T#10S,
		tDoorClose := T#10S,
		tHatchUnlock := T#5S,
		tChuckOpen := T#10S,
		tChuckClose := T#10S,
		tCycleStart := T#10S
	); // Штатные пределы ожидания технологических подтверждений станков
	stAxisTimeouts : ST_AXIS_TIMEOUTS := (
		xDisableOnError := TRUE,
		tPowerFeedbackLossTimeout := T#500MS,
		tPowerTimeout := T#5S,
		tResetTimeout := T#5S,
		tStopTimeout := T#5S,
		tHomeTimeout := T#30S,
		tMoveTimeout := T#15S
	); // Общий профиль ожиданий для осей X/Y/Z
	stAxisGroupTimeouts : ST_AXIS_GROUP_TIMEOUTS := (
		tPowerTimeout := T#5S,
		tGroupTimeout := T#5S,
		tStopTimeout := T#5S,
		tHaltTimeout := T#5S,
		tHomeTimeout := T#30S,
		tMoveTimeout := T#30S
	); // Ожидания координатной группы XYZ
	tPointCheckStartTimeout : TIME := T#2S; // Ожидание фактического старта проверки точки
	tSimulationDynamicsTimeout : TIME := T#60S; // Stop -> Disable -> Dynamic Limits -> Enable
	tHmiWatchdogTimeout : TIME := T#2S; // Потеря основного heartbeat HMI
	tMobileMotionWatchdogTimeout : TIME := T#2S; // Потеря heartbeat мобильного движения
	tPointCheckWatchdogTimeout : TIME := T#2S; // Потеря владельца проверки точки
	tHmiCommandFreshnessTimeout : TIME := T#3S; // Максимальный возраст подтверждаемой команды HMI

	//Порядок команд для смены, загрузки и выгрузки станков
	CHANGE_MACHINE : ARRAY [0..40] OF ST_MACHINE_RECIPE // Рецепт смены детали в станке
	:=[
	   (eCommand := E_MACHINE_STATE.DOOR_OPEN),
	   (eCommand := E_MACHINE_STATE.ROBOT_ACTION, eRobotAction := E_ROBOT_ACTION.ROTATE_TO_DETAIL),
	   (eCommand := E_MACHINE_STATE.ROBOT_ACTION, eRobotAction := E_ROBOT_ACTION.UNCLAMP_2),
	   (eCommand := E_MACHINE_STATE.ROBOT_MOVE, stPoint := E_MACHINE_POINTS.CHUCK_APPROACH),
	   (eCommand := E_MACHINE_STATE.ROBOT_MOVE, stPoint := E_MACHINE_POINTS.CHUCK),
	   (eCommand := E_MACHINE_STATE.ROBOT_ACTION, eRobotAction := E_ROBOT_ACTION.CLAMP_2),
	   (eCommand := E_MACHINE_STATE.CHUCK_OPEN),
	   (eCommand := E_MACHINE_STATE.ROBOT_MOVE, stPoint := E_MACHINE_POINTS.CHUCK_APPROACH),
	   (eCommand := E_MACHINE_STATE.ROBOT_ACTION, eRobotAction := E_ROBOT_ACTION.ROTATE_TO_BLANK),
	   (eCommand := E_MACHINE_STATE.ROBOT_MOVE, stPoint := E_MACHINE_POINTS.CHUCK),
	   (eCommand := E_MACHINE_STATE.CHUCK_CLOSE),
	   (eCommand := E_MACHINE_STATE.ROBOT_ACTION, eRobotAction := E_ROBOT_ACTION.UNCLAMP_1),
	   (eCommand := E_MACHINE_STATE.ROBOT_MOVE, stPoint := E_MACHINE_POINTS.CHUCK_APPROACH),
	   (eCommand := E_MACHINE_STATE.ROBOT_MOVE, stPoint := E_MACHINE_POINTS.ABOVE, xRobotDone := TRUE),
	   (eCommand := E_MACHINE_STATE.DOOR_CLOSE),
	   (eCommand := E_MACHINE_STATE.CYCLE_START),
	   (eCommand := E_MACHINE_STATE.DONE)
	   
	   
	   
	   
];
	LOAD_MACHINE : ARRAY [0..40] OF ST_MACHINE_RECIPE // Рецепт загрузки станка
	:=[
	   (eCommand := E_MACHINE_STATE.DOOR_OPEN),
	   (eCommand := E_MACHINE_STATE.ROBOT_ACTION, eRobotAction := E_ROBOT_ACTION.ROTATE_TO_BLANK),
	   (eCommand := E_MACHINE_STATE.ROBOT_MOVE, stPoint := E_MACHINE_POINTS.CHUCK_APPROACH),
	   (eCommand := E_MACHINE_STATE.ROBOT_MOVE, stPoint := E_MACHINE_POINTS.CHUCK),
	   (eCommand := E_MACHINE_STATE.CHUCK_CLOSE),
	   (eCommand := E_MACHINE_STATE.ROBOT_ACTION, eRobotAction := E_ROBOT_ACTION.UNCLAMP_1),
	   (eCommand := E_MACHINE_STATE.ROBOT_MOVE, stPoint := E_MACHINE_POINTS.CHUCK_APPROACH),
	   (eCommand := E_MACHINE_STATE.ROBOT_MOVE, stPoint := E_MACHINE_POINTS.ABOVE, xRobotDone := TRUE),
	   (eCommand := E_MACHINE_STATE.DOOR_CLOSE),
	   (eCommand := E_MACHINE_STATE.CYCLE_START),
	   (eCommand := E_MACHINE_STATE.DONE)
	];

	UNLOAD_MACHINE : ARRAY [0..40] OF ST_MACHINE_RECIPE // Рецепт выгрузки станка
	:=[
	   (eCommand := E_MACHINE_STATE.DOOR_OPEN),
	   (eCommand := E_MACHINE_STATE.ROBOT_ACTION, eRobotAction := E_ROBOT_ACTION.ROTATE_TO_DETAIL),
	   (eCommand := E_MACHINE_STATE.ROBOT_ACTION, eRobotAction := E_ROBOT_ACTION.UNCLAMP_2),
	   (eCommand := E_MACHINE_STATE.ROBOT_MOVE, stPoint := E_MACHINE_POINTS.CHUCK_APPROACH),
	   (eCommand := E_MACHINE_STATE.ROBOT_MOVE, stPoint := E_MACHINE_POINTS.CHUCK),
	   (eCommand := E_MACHINE_STATE.ROBOT_ACTION, eRobotAction := E_ROBOT_ACTION.CLAMP_2),
	   (eCommand := E_MACHINE_STATE.CHUCK_OPEN),
	   (eCommand := E_MACHINE_STATE.ROBOT_MOVE, stPoint := E_MACHINE_POINTS.CHUCK_APPROACH),
	   (eCommand := E_MACHINE_STATE.ROBOT_MOVE, stPoint := E_MACHINE_POINTS.ABOVE, xRobotDone := TRUE),
	   (eCommand := E_MACHINE_STATE.DOOR_CLOSE),
	   (eCommand := E_MACHINE_STATE.DONE)
	];
END_VAR

// Device/Application/GVL/GVL_DETAIL
{attribute 'qualified_only'}
VAR_GLOBAL
	astMagazine : ARRAY [1..GVL_CELL_SETTINGS.MagazineCount] OF ST_MAGAZINE_INVENTORY; // Три зоны двух магазинов
END_VAR

// Device/Application/GVL/GVL_AXIS
{attribute 'qualified_only'}
VAR_GLOBAL
	arrAxis : ARRAY [1..3] OF ST_AXIS; // Команды, статусы и диагностика осей X, Y, Z
END_VAR

// Device/Application/GVL/GVL_MULTI_TYPE
{attribute 'qualified_only'}
VAR_GLOBAL
	Config       : ST_MULTI_TYPE_CONFIG; // Активная конфигурация типов продукции
	ConfigStatus : ST_MULTI_TYPE_CONFIG_STATUS; // Разрешения редактирования конфигурации
	CycleStatus  : ST_CELL_CYCLE_STATUS; // Диагностика универсального автомата ячейки
END_VAR

// Device/Application/GVL/GVL_MOTION_MANAGER
{attribute 'qualified_only'}
VAR_GLOBAL
	stMotionManager : ST_MOTION_MANAGER; // Команды, статусы и диагностика менеджера движения
END_VAR

// Device/Application/GVL/GVL_PHYSICAL_IO
{attribute 'qualified_only'}
VAR_GLOBAL
	// Привязать существующие BOOL через Device I/O Mapping. Адреса ниже —
	// проект фиксированного процесса с базой байта 256, НЕ адреса по умолчанию MC522.
	// Не добавлять AT поверх Device I/O Mapping: у выхода должен быть один писатель.
	// MC522 16 DI/16 DO + 5×GL200-DI16 + 2×GL200-DQ16D; 84 BOOL DI, 2 HSC и 47 DO.
	xMappingVerified : BOOL := FALSE; // Наладчик подтверждает после полной проверки клемм; не RETAIN
	xNormalActive : BOOL; // NORMAL и подтверждённая карта были применены перед RunSafety
	stGripperFeedback : ST_GRIPPER_STATUS;
	stGripperCommand : ST_GRIPPER_COMMAND;
	axMachineHatchClose : ARRAY [1..3] OF BOOL; // Удерживаемые уровни однокатушечных люков
	axGkPartAtEnd : ARRAY [1..2] OF BOOL; // Фильтрованная фиксация ГК 1/2: NORMAL с проверенной картой либо разрешённой подменой DI
	xDiMachine1Ready : BOOL; // %IX256.2; MC522: DI_CH2; Станок готов к работе с роботом. 1 — указанное состояние; 1→0 без задержки
	xDiMachine1Alarm : BOOL; // %IX256.3; MC522: DI_CH3; Авария станка. 1 — авария; снимается физически человеком; 0→1 без задержки
	xDiMachine1DoorOpen : BOOL; // %IX256.4; MC522: DI_CH4; Роботный люк открыт. 1 — указанное состояние; 1→0 без задержки
	xDiMachine1DoorClosed : BOOL; // %IX256.5; MC522: DI_CH5; Роботный люк закрыт. 1 — указанное состояние; 1→0 без задержки
	xDiMachine1HatchLocked : BOOL; // %IX256.6; MC522: DI_CH6; Замок роботного люка заперт. 1 — замок люка заперт; 0 — запирание не подтверждено; 1→0 без задержки
	xDiMachine1SafetyDoorOpen : BOOL; // %IX256.7; MC522: DI_CH7; Операторская дверь открыта. 1 — указанное состояние; 1→0 без задержки
	xDiMachine1SafetyDoorClosed : BOOL; // %IX257.0; MC522: DI_CH8; Операторская дверь закрыта. 1 — указанное состояние; 1→0 без задержки
	xDiMachine1ChuckClamped : BOOL; // %IX257.1; MC522: DI_CH9; Патрон зажат. 1 — указанное состояние; 1→0 без задержки
	xDiMachine1ChuckUnclamped : BOOL; // %IX257.2; MC522: DI_CH10; Патрон разжат. 1 — указанное состояние; 1→0 без задержки
	xDiMachine1CycleActive : BOOL; // %IX257.3; MC522: DI_CH11; Цикл обработки активен. 1 — указанное состояние
	xDiMachine1CycleDone : BOOL; // %IX257.4; MC522: DI_CH12; Цикл обработки завершён. 1 — указанное состояние
	xDiMachine2Ready : BOOL; // %IX257.5; MC522: DI_CH13; Станок готов к работе с роботом. 1 — указанное состояние; 1→0 без задержки
	xDiMachine2Alarm : BOOL; // %IX257.6; MC522: DI_CH14; Авария станка. 1 — авария; снимается физически человеком; 0→1 без задержки
	xDiMachine2DoorOpen : BOOL; // %IX257.7; MC522: DI_CH15; Роботный люк открыт. 1 — указанное состояние; 1→0 без задержки
	xDiMachine2DoorClosed : BOOL; // %IX258.0; GL200-DI16 #1: CH0; Роботный люк закрыт. 1 — указанное состояние; 1→0 без задержки
	xDiMachine2HatchLocked : BOOL; // %IX258.1; GL200-DI16 #1: CH1; Замок роботного люка заперт. 1 — замок люка заперт; 0 — запирание не подтверждено; 1→0 без задержки
	xDiMachine2SafetyDoorOpen : BOOL; // %IX258.2; GL200-DI16 #1: CH2; Операторская дверь открыта. 1 — указанное состояние; 1→0 без задержки
	xDiMachine2SafetyDoorClosed : BOOL; // %IX258.3; GL200-DI16 #1: CH3; Операторская дверь закрыта. 1 — указанное состояние; 1→0 без задержки
	xDiMachine2ChuckClamped : BOOL; // %IX258.4; GL200-DI16 #1: CH4; Патрон зажат. 1 — указанное состояние; 1→0 без задержки
	xDiMachine2ChuckUnclamped : BOOL; // %IX258.5; GL200-DI16 #1: CH5; Патрон разжат. 1 — указанное состояние; 1→0 без задержки
	xDiMachine2CycleActive : BOOL; // %IX258.6; GL200-DI16 #1: CH6; Цикл обработки активен. 1 — указанное состояние
	xDiMachine2CycleDone : BOOL; // %IX258.7; GL200-DI16 #1: CH7; Цикл обработки завершён. 1 — указанное состояние
	xDiMachine3Ready : BOOL; // %IX259.0; GL200-DI16 #1: CH8; Станок готов к работе с роботом. 1 — указанное состояние; 1→0 без задержки
	xDiMachine3Alarm : BOOL; // %IX259.1; GL200-DI16 #1: CH9; Авария станка. 1 — авария; снимается физически человеком; 0→1 без задержки
	xDiMachine3DoorOpen : BOOL; // %IX259.2; GL200-DI16 #1: CH10; Роботный люк открыт. 1 — указанное состояние; 1→0 без задержки
	xDiMachine3DoorClosed : BOOL; // %IX259.3; GL200-DI16 #1: CH11; Роботный люк закрыт. 1 — указанное состояние; 1→0 без задержки
	xDiMachine3HatchLocked : BOOL; // %IX259.4; GL200-DI16 #1: CH12; Замок роботного люка заперт. 1 — замок люка заперт; 0 — запирание не подтверждено; 1→0 без задержки
	xDiMachine3SafetyDoorOpen : BOOL; // %IX259.5; GL200-DI16 #1: CH13; Операторская дверь открыта. 1 — указанное состояние; 1→0 без задержки
	xDiMachine3SafetyDoorClosed : BOOL; // %IX259.6; GL200-DI16 #1: CH14; Операторская дверь закрыта. 1 — указанное состояние; 1→0 без задержки
	xDiMachine3ChuckClamped : BOOL; // %IX259.7; GL200-DI16 #1: CH15; Патрон зажат. 1 — указанное состояние; 1→0 без задержки
	xDiMachine3ChuckUnclamped : BOOL; // %IX260.0; GL200-DI16 #2: CH0; Патрон разжат. 1 — указанное состояние; 1→0 без задержки
	xDiMachine3CycleActive : BOOL; // %IX260.1; GL200-DI16 #2: CH1; Цикл обработки активен. 1 — указанное состояние
	xDiMachine3CycleDone : BOOL; // %IX260.2; GL200-DI16 #2: CH2; Цикл обработки завершён. 1 — указанное состояние
	xDiGripper1Open : BOOL; // %IX260.3; GL200-DI16 #2: CH3; Захват 1 открыт. 1 — указанная позиция; в Modbus источником остаётся SC-500; 1→0 без задержки
	xDiGripper1Closed : BOOL; // %IX260.4; GL200-DI16 #2: CH4; Захват 1 закрыт. 1 — указанная позиция; в Modbus источником остаётся SC-500; 1→0 без задержки
	xDiGripper2Open : BOOL; // %IX260.5; GL200-DI16 #2: CH5; Захват 2 открыт. 1 — указанная позиция; в Modbus источником остаётся SC-500; 1→0 без задержки
	xDiGripper2Closed : BOOL; // %IX260.6; GL200-DI16 #2: CH6; Захват 2 закрыт. 1 — указанная позиция; в Modbus источником остаётся SC-500; 1→0 без задержки
	xDiRotatedToBlank : BOOL; // %IX260.7; GL200-DI16 #2: CH7; Поворот к заготовке. 1 — указанная позиция; в Modbus источником остаётся SC-500; 1→0 без задержки
	xDiRotatedToDetail : BOOL; // %IX261.0; GL200-DI16 #2: CH8; Поворот к детали. 1 — указанная позиция; в Modbus источником остаётся SC-500; 1→0 без задержки
	xDiCellStartButtonInput : BOOL; // %IX261.1; GL200-DI16 #2: CH9; Запустить ячейку в работу. 1 — кнопка пуска нажата
	xDiCellStopButtonInput : BOOL; // %IX261.2; GL200-DI16 #2: CH10; Вывести ячейку из работы. 1 — кнопка останова нажата; 0→1 без задержки
	xDiCellResetButtonInput : BOOL; // %IX261.3; GL200-DI16 #2: CH11; Сбросить ошибки ячейку. 1 — кнопка нажата; локальный сброс программных ошибок ячейки, без сброса физической аварии станка
	xDiEmergencyStopStation1Ok : BOOL; // %IX261.4; GL200-DI16 #2: CH12; Аварийный грибок 1. Физический xDi: 1 — грибок отжат, 0 — нажат/обрыв; программный xEmergency: TRUE — нажат; потеря физической 1 проходит без задержки
	xDiEmergencyStopStation2Ok : BOOL; // %IX261.5; GL200-DI16 #2: CH13; Аварийный грибок 2. Физический xDi: 1 — грибок отжат, 0 — нажат/обрыв; программный xEmergency: TRUE — нажат; потеря физической 1 проходит без задержки
	xDiEmergencyStopStation3Ok : BOOL; // %IX261.6; GL200-DI16 #2: CH14; Аварийный грибок 3. Физический xDi: 1 — грибок отжат, 0 — нажат/обрыв; программный xEmergency: TRUE — нажат; потеря физической 1 проходит без задержки
	xDiEmergencyStopStation4Ok : BOOL; // %IX261.7; GL200-DI16 #2: CH15; Аварийный грибок 4. Физический xDi: 1 — грибок отжат, 0 — нажат/обрыв; программный xEmergency: TRUE — нажат; потеря физической 1 проходит без задержки
	xDiEmergencyStopCabinet1Ok : BOOL; // %IX262.0; GL200-DI16 #3: CH0; Аварийный грибок 5. Физический xDi: 1 — грибок отжат, 0 — нажат/обрыв; программный xEmergency: TRUE — нажат; потеря физической 1 проходит без задержки
	xDiEmergencyStopCabinet2Ok : BOOL; // %IX262.1; GL200-DI16 #3: CH1; Аварийный грибок 6. Физический xDi: 1 — грибок отжат, 0 — нажат/обрыв; программный xEmergency: TRUE — нажат; потеря физической 1 проходит без задержки
	xDiEmergencyStopMpgOk : BOOL; // %IX262.2; GL200-DI16 #3: CH2; Аварийный грибок 7. Физический xDi: 1 — грибок отжат, 0 — нажат/обрыв; программный xEmergency: TRUE — нажат; потеря физической 1 проходит без задержки
	xDiDoor1LockClosed : BOOL; // %IX262.3; GL200-DI16 #3: CH3; Замок двери 1 закрыт. 1 — замок закрыт; 0 — закрытие не подтверждено; 1→0 без задержки
	xDiDoor2LockClosed : BOOL; // %IX262.4; GL200-DI16 #3: CH4; Замок двери 2 закрыт. 1 — замок закрыт; 0 — закрытие не подтверждено; 1→0 без задержки
	xDiDoor3LockClosed : BOOL; // %IX262.5; GL200-DI16 #3: CH5; Замок двери 3 закрыт. 1 — замок закрыт; 0 — закрытие не подтверждено; 1→0 без задержки
	xDiDoor4LockClosed : BOOL; // %IX262.6; GL200-DI16 #3: CH6; Замок двери 4 закрыт. 1 — замок закрыт; 0 — закрытие не подтверждено; 1→0 без задержки
	xDiSafetyRelayOkInput : BOOL; // %IX262.7; GL200-DI16 #3: CH7; Реле безопасности 1, взведено. 1 — норма; потеря нормы проходит без задержки; 1→0 без задержки
	xDiPhaseRelayOkInput : BOOL; // %IX263.0; GL200-DI16 #3: CH8; Фазы совпадают. 1 — норма; потеря нормы проходит без задержки; 1→0 без задержки
	xDiPressureRelayOkInput : BOOL; // %IX263.1; GL200-DI16 #3: CH9; Давление стабильно. 1 — норма; потеря нормы проходит без задержки; 1→0 без задержки
	xDiMpgAxisXInput : BOOL; // %IX263.2; GL200-DI16 #3: CH10; Выбор оси X. 1 — выбрана ось X
	xDiMpgAxisYInput : BOOL; // %IX263.3; GL200-DI16 #3: CH11; Выбор оси Y. 1 — выбрана ось Y
	xDiMpgAxisZInput : BOOL; // %IX263.4; GL200-DI16 #3: CH12; Выбор оси Z. 1 — выбрана ось Z
	xDiMpgMultiplier1Input : BOOL; // %IX263.5; GL200-DI16 #3: CH13; Множитель ×1. 1 — выбран множитель ×1
	xDiMpgMultiplier10Input : BOOL; // %IX263.6; GL200-DI16 #3: CH14; Множитель ×10. 1 — выбран множитель ×10
	xDiMpgMultiplier100Input : BOOL; // %IX263.7; GL200-DI16 #3: CH15; Множитель ×100. 1 — выбран множитель ×100
	xDiMagazine1LockIn : BOOL; // %IX264.0; GL200-DI16 #4: CH0; Замок втянут. 1 — геркон сработал; 1→0 без задержки
	xDiMagazine1LockOut : BOOL; // %IX264.1; GL200-DI16 #4: CH1; Замок выдвинут. 1 — геркон сработал; 1→0 без задержки
	xDiMagazine1StopIn : BOOL; // %IX264.2; GL200-DI16 #4: CH2; Фиксатор выдвинут. 1 — геркон сработал; 1→0 без задержки
	xDiMagazine1StopOut : BOOL; // %IX264.3; GL200-DI16 #4: CH3; Фиксатор втянут. 1 — геркон сработал; 1→0 без задержки
	xDiMagazine1LiftUp : BOOL; // %IX264.4; GL200-DI16 #4: CH4; Подъёмник вверху. 1 — геркон сработал; 1→0 без задержки
	xDiMagazine1LiftDown : BOOL; // %IX264.5; GL200-DI16 #4: CH5; Подъёмник внизу. 1 — геркон сработал; 1→0 без задержки
	xDiDoor1UnlockButton : BOOL; // %IX265.4; GL200-DI16 #4: CH12; Кнопка запроса открытия двери 1. 1 — нажата
	xDiDoor2UnlockButton : BOOL; // %IX265.5; GL200-DI16 #4: CH13; Кнопка запроса открытия двери 2. 1 — нажата
	xDiDoor3UnlockButton : BOOL; // %IX265.6; GL200-DI16 #4: CH14; Кнопка запроса открытия двери 3. 1 — нажата
	xDiDoor4UnlockButton : BOOL; // %IX265.7; GL200-DI16 #4: CH15; Кнопка запроса открытия двери 4. 1 — нажата
	xDiGk1DriveAlarm : BOOL; // %IX264.6; GL200-DI16 #4: CH6; ГК привод — Авария. 1 — авария частотника конвейера ГК. В NORMAL используется FB_GEOMETRY_CONTROL без задержки.
	xDiGk1DriveRunning : BOOL; // %IX264.7; GL200-DI16 #4: CH7; ГК привод — Работа. 1 — привод конвейера ГК в работе. В NORMAL используется FB_GEOMETRY_CONTROL без задержки.
	xDiGk1PartAtEnd : BOOL; // %IX265.0; GL200-DI16 #4: CH8; Датчик фиксации детали на конце конвейера. 1 — деталь на конце конвейера ГК. Передний фронт фильтруется; потеря уровня сразу, изъятие подтверждается FB_GEOMETRY_CONTROL через 3 секунды.
	xDiGk2DriveAlarm : BOOL; // %IX265.1; GL200-DI16 #4: CH9; ГК привод — Авария. 1 — авария частотника конвейера ГК. В NORMAL используется FB_GEOMETRY_CONTROL без задержки.
	xDiGk2DriveRunning : BOOL; // %IX265.2; GL200-DI16 #4: CH10; ГК привод — Работа. 1 — привод конвейера ГК в работе. В NORMAL используется FB_GEOMETRY_CONTROL без задержки.
	xDiGk2PartAtEnd : BOOL; // %IX265.3; GL200-DI16 #4: CH11; Датчик фиксации детали на конце конвейера. 1 — деталь на конце конвейера ГК. Передний фронт фильтруется; потеря уровня сразу, изъятие подтверждается FB_GEOMETRY_CONTROL через 3 секунды.
	xDiMagazine2LockIn : BOOL; // %IX266.0; GL200-DI16 #5: CH0; Замок втянут. 1 — геркон сработал; 1→0 без задержки
	xDiMagazine2LockOut : BOOL; // %IX266.1; GL200-DI16 #5: CH1; Замок выдвинут. 1 — геркон сработал; 1→0 без задержки
	xDiMagazine2StopIn : BOOL; // %IX266.2; GL200-DI16 #5: CH2; Фиксатор выдвинут. 1 — геркон сработал; 1→0 без задержки
	xDiMagazine2StopOut : BOOL; // %IX266.3; GL200-DI16 #5: CH3; Фиксатор втянут. 1 — геркон сработал; 1→0 без задержки
	xDiMagazine2LiftUp : BOOL; // %IX266.4; GL200-DI16 #5: CH4; Подъёмник вверху. 1 — геркон сработал; 1→0 без задержки
	xDiMagazine2LiftDown : BOOL; // %IX266.5; GL200-DI16 #5: CH5; Подъёмник внизу. 1 — геркон сработал; 1→0 без задержки
	xDoMachine1HatchClosed : BOOL; // %QX256.0; MC522: DO_CH0; Открыть роботный люк/Закрыть роботный люк. 0 — открыть люк; 1 — закрыть. Уровень удерживается между командами.
	xDoMachine1HatchUnLock : BOOL; // %QX256.1; MC522: DO_CH1; Открыть замок люка. 1 — команда активна
	xDoMachine1ClampChuck : BOOL; // %QX256.2; MC522: DO_CH2; Зажать патрон. 1 — команда активна
	xDoMachine1UnclampChuck : BOOL; // %QX256.3; MC522: DO_CH3; Разжать патрон. 1 — команда активна
	xDoMachine1StartCycle : BOOL; // %QX256.4; MC522: DO_CH4; Запустить обработку. 1 — запуск обработки; штатно — команда FB станка; прямой ручной I/O удерживает выбранный уровень
	xDoMachine2HatchClosed : BOOL; // %QX256.5; MC522: DO_CH5; Открыть роботный люк/Закрыть роботный люк. 0 — открыть люк; 1 — закрыть. Уровень удерживается между командами.
	xDoMachine2HatchUnLock : BOOL; // %QX256.6; MC522: DO_CH6; Открыть замок люка. 1 — команда активна
	xDoMachine2ClampChuck : BOOL; // %QX256.7; MC522: DO_CH7; Зажать патрон. 1 — команда активна
	xDoMachine2UnclampChuck : BOOL; // %QX257.0; MC522: DO_CH8; Разжать патрон. 1 — команда активна
	xDoMachine2StartCycle : BOOL; // %QX257.1; MC522: DO_CH9; Запустить обработку. 1 — запуск обработки; штатно — команда FB станка; прямой ручной I/O удерживает выбранный уровень
	xDoMachine3HatchClosed : BOOL; // %QX257.2; MC522: DO_CH10; Открыть роботный люк/Закрыть роботный люк. 0 — открыть люк; 1 — закрыть. Уровень удерживается между командами.
	xDoMachine3HatchUnLock : BOOL; // %QX257.3; MC522: DO_CH11; Открыть замок люка. 1 — команда активна
	xDoMachine3ClampChuck : BOOL; // %QX257.4; MC522: DO_CH12; Зажать патрон. 1 — команда активна
	xDoMachine3UnclampChuck : BOOL; // %QX257.5; MC522: DO_CH13; Разжать патрон. 1 — команда активна
	xDoMachine3StartCycle : BOOL; // %QX257.6; MC522: DO_CH14; Запустить обработку. 1 — запуск обработки; штатно — команда FB станка; прямой ручной I/O удерживает выбранный уровень
	xDoGripper1Open : BOOL; // %QX257.7; MC522: DO_CH15; Открыть захват 1 / Закрыть захват 1. 0 — закрыть; 1 — открыть. Штатное управление физическим DO — SoftMotion NORMAL; прямой ручной I/O задаёт уровень независимо от режима привода
	xDoGripper2Open : BOOL; // %QX258.0; GL200-DQ16D #1: CH0; Открыть захват 2 / Закрыть захват 2. 0 — закрыть; 1 — открыть. Штатное управление физическим DO — SoftMotion NORMAL; прямой ручной I/O задаёт уровень независимо от режима привода
	xDoRotateToDetail : BOOL; // %QX258.1; GL200-DQ16D #1: CH1; Повернуть к заготовке / Повернуть к детали. 0 — к заготовке; 1 — к детали. Штатное управление физическим DO — SoftMotion NORMAL; прямой ручной I/O задаёт уровень независимо от режима привода
	xDoDoor1Unlock : BOOL; // %QX258.2; GL200-DQ16D #1: CH2; Открыть замок двери 1. 1 — разблокировать замок двери
	xDoDoor2Unlock : BOOL; // %QX258.3; GL200-DQ16D #1: CH3; Открыть замок двери 2. 1 — разблокировать замок двери
	xDoDoor3Unlock : BOOL; // %QX258.4; GL200-DQ16D #1: CH4; Открыть замок двери 3. 1 — разблокировать замок двери
	xDoDoor4Unlock : BOOL; // %QX258.5; GL200-DQ16D #1: CH5; Открыть замок двери 4. 1 — разблокировать замок двери
	xDoSafetyRelayReset : BOOL; // %QX258.6; GL200-DQ16D #1: CH6; Сигнал сброса на реле безопасности 1. Штатно — импульс сброса реле безопасности, без сброса физической аварии станка; прямой ручной I/O удерживает выбранный уровень
	xDoSignalTowerGreenOutput : BOOL; // %QX258.7; GL200-DQ16D #1: CH7; Зеленый цвет. Уровень с миганием из PLC_PRG.RunSignalTower
	xDoSignalTowerAmberOutput : BOOL; // %QX259.0; GL200-DQ16D #1: CH8; Желтый цвет. Уровень с миганием из PLC_PRG.RunSignalTower
	xDoSignalTowerRedOutput : BOOL; // %QX259.1; GL200-DQ16D #1: CH9; Красный цвет. Уровень с миганием из PLC_PRG.RunSignalTower
	xDoDoor1ButtonLamp : BOOL; // %QX259.3; GL200-DQ16D #1: CH11; Световая индикация кнопки 1. Готовый уровень индикации из FB_CELL_SAFETY
	xDoDoor2ButtonLamp : BOOL; // %QX259.4; GL200-DQ16D #1: CH12; Световая индикация кнопки 2. Готовый уровень индикации из FB_CELL_SAFETY
	xDoDoor3ButtonLamp : BOOL; // %QX259.5; GL200-DQ16D #1: CH13; Световая индикация кнопки 3. Готовый уровень индикации из FB_CELL_SAFETY
	xDoDoor4ButtonLamp : BOOL; // %QX259.6; GL200-DQ16D #1: CH14; Световая индикация кнопки 4. Готовый уровень индикации из FB_CELL_SAFETY
	xDoMagazine1LockIn : BOOL; // %QX259.7; GL200-DQ16D #1: CH15; Замок втянут (катушка). 1 — катушка включена; штатная логика исключает встречные катушки; в прямом ручном I/O этого ограничения нет
	xDoMagazine1LockOut : BOOL; // %QX260.0; GL200-DQ16D #2: CH0; Замок выдвинут (катушка). 1 — катушка включена; штатная логика исключает встречные катушки; в прямом ручном I/O этого ограничения нет
	xDoMagazine1StopIn : BOOL; // %QX260.1; GL200-DQ16D #2: CH1; Фиксатор выдвинут (катушка). 1 — катушка включена; штатная логика исключает встречные катушки; в прямом ручном I/O этого ограничения нет
	xDoMagazine1StopOut : BOOL; // %QX260.2; GL200-DQ16D #2: CH2; Фиксатор втянут (катушка). 1 — катушка включена; штатная логика исключает встречные катушки; в прямом ручном I/O этого ограничения нет
	xDoMagazine1LiftUp : BOOL; // %QX260.3; GL200-DQ16D #2: CH3; Подъёмник вверху (катушка). 1 — катушка включена; штатная логика исключает встречные катушки; в прямом ручном I/O этого ограничения нет
	xDoMagazine1LiftDown : BOOL; // %QX260.4; GL200-DQ16D #2: CH4; Подъёмник внизу (катушка). 1 — катушка включена; штатная логика исключает встречные катушки; в прямом ручном I/O этого ограничения нет
	xDoCellAlarmHorn : BOOL; // %QX259.2; GL200-DQ16D #1: CH10; Гудок. Штатно — звук при новой аварии: 0–60 с, по умолчанию 2 с; 0 отключает автоматический звук. Прямой ручной I/O удерживает выбранный уровень
	xDoGk1DriveRun : BOOL; // %QX260.5; GL200-DQ16D #2: CH5; ГК привод — Пуск / Стоп. 1 — пуск, 0 — стоп. Штатный владелец FB_GEOMETRY_CONTROL; в прямом ручном I/O уровень задаётся вручную.
	xDoGk1DriveReset : BOOL; // %QX260.6; GL200-DQ16D #2: CH6; ГК привод — Сброс аварии. Импульс сброса частотника от FB_GEOMETRY_CONTROL; длительность задаётся в таймаутах ячейки.
	xDoMagazine2LockIn : BOOL; // %QX261.1; GL200-DQ16D #2: CH9; Замок втянут (катушка). 1 — катушка включена; штатная логика исключает встречные катушки; в прямом ручном I/O этого ограничения нет
	xDoMagazine2LockOut : BOOL; // %QX261.2; GL200-DQ16D #2: CH10; Замок выдвинут (катушка). 1 — катушка включена; штатная логика исключает встречные катушки; в прямом ручном I/O этого ограничения нет
	xDoMagazine2StopIn : BOOL; // %QX261.3; GL200-DQ16D #2: CH11; Фиксатор выдвинут (катушка). 1 — катушка включена; штатная логика исключает встречные катушки; в прямом ручном I/O этого ограничения нет
	xDoMagazine2StopOut : BOOL; // %QX261.4; GL200-DQ16D #2: CH12; Фиксатор втянут (катушка). 1 — катушка включена; штатная логика исключает встречные катушки; в прямом ручном I/O этого ограничения нет
	xDoMagazine2LiftUp : BOOL; // %QX261.5; GL200-DQ16D #2: CH13; Подъёмник вверху (катушка). 1 — катушка включена; штатная логика исключает встречные катушки; в прямом ручном I/O этого ограничения нет
	xDoMagazine2LiftDown : BOOL; // %QX261.6; GL200-DQ16D #2: CH14; Подъёмник внизу (катушка). 1 — катушка включена; штатная логика исключает встречные катушки; в прямом ручном I/O этого ограничения нет
	xDoGk2DriveRun : BOOL; // %QX260.7; GL200-DQ16D #2: CH7; ГК привод — Пуск / Стоп. 1 — пуск, 0 — стоп. Штатный владелец FB_GEOMETRY_CONTROL; в прямом ручном I/O уровень задаётся вручную.
	xDoGk2DriveReset : BOOL; // %QX261.0; GL200-DQ16D #2: CH8; ГК привод — Сброс аварии. Импульс сброса частотника от FB_GEOMETRY_CONTROL; длительность задаётся в таймаутах ячейки.
END_VAR

// Device/Application/GVL/GVL_TWO_PALLET
{attribute 'qualified_only'}
VAR_GLOBAL
	Axis1 : REFERENCE TO AXIS_REF_SM3; // Каждый скан REF= Magazine_1 в RunTwoPalletAxis
	Axis2 : REFERENCE TO AXIS_REF_SM3; // Каждый скан REF= Magazine_2 в RunTwoPalletAxis
	astAxis : ARRAY [1..2] OF ST_AXIS;
	astInput : ARRAY [1..2] OF ST_TWO_PALLET_INPUT; // Физические входы: НЕ записываются из HMI
	astOutput : ARRAY [1..2] OF ST_TWO_PALLET_OUTPUT;
	astSimulationConfig : ARRAY [1..2] OF ST_TWO_PALLET_CONFIG; // Только виртуальная среда; не RETAIN
	astActiveConfig : ARRAY [1..2] OF ST_TWO_PALLET_CONFIG; // Конфигурация текущей среды
	astStatus : ARRAY [1..2] OF ST_TWO_PALLET_STATUS;
	astDiag : ARRAY [1..2] OF ST_TWO_PALLET_DIAG;
	astError : ARRAY [1..2] OF ST_TWO_PALLET_ERRORS;
	auiCommand : ARRAY [1..2] OF UINT;
	auiValue : ARRAY [1..2] OF UINT;
	audiRevision : ARRAY [1..2] OF UDINT;
	xModeChangeAllowed : BOOL;
	xModeChanged : BOOL;
	astStatic : ARRAY [1..2] OF ST_MAGAZINE_INVENTORY;
	axSimulationAutoSwapEnabled : ARRAY [1..2] OF BOOL; // Только виртуальная среда; не RETAIN
END_VAR
VAR_GLOBAL RETAIN
	uiMode : UINT := UINT#1; // По умолчанию два двухпалетных; 0: два статичных; 1: два двухпалетных
	astConfig : ARRAY [1..2] OF ST_TWO_PALLET_CONFIG;
	astStore : ARRAY [1..2] OF ST_TWO_PALLET_STORE;
	axAutoSwapEnabled : ARRAY [1..2] OF BOOL := [TRUE, TRUE];
	xAutoSwapDefaultsApplied : BOOL; // Однократная инициализация новой RETAIN-настройки
END_VAR

VAR_GLOBAL PERSISTENT RETAIN
	// Постоянный шаг сетки для расчёта координат робота, отдельно по типам магазинов.
	lrStaticPitchX : LREAL := 60.0;
	lrStaticPitchY : LREAL := 60.0;
	lrTwinPitchX : LREAL := 70.0;
	lrTwinPitchY : LREAL := 70.0;
END_VAR

// Device/Application/PLC_PRG
PROGRAM PLC_PRG
VAR
	GEOMETRY : ARRAY [1..2] OF FB_GEOMETRY_CONTROL;
	GEOMETRY_SIM : ARRAY [1..2] OF FB_GEOMETRY_CONTROL_SIMULATION;
	xGeometryInitialized : BOOL;
	xGeometryEnvironmentChanged : BOOL;
	eGeometryPreviousEnvironment : E_CELL_TEST_ENVIRONMENT;
	uiGeometry : UINT;
	uiGeometryMachine : UINT;
	uiGeometryDi : UINT;
	udiGeometryRequest : UDINT;
	stGeometryRequest : ST_GEOMETRY_REQUEST;
	stGeometryConfig : ST_GEOMETRY_CONFIG;
	stGeometryCall : ST_GEOMETRY_CALL;
	stGeometryEmptyCall : ST_GEOMETRY_CALL;
	xGeometryConfigValid : BOOL;
	xGeometryDriveAlarm : BOOL;
	xGeometryDriveRunning : BOOL;
	xGeometryPartAtEnd : BOOL;
	stGeometrySignals : ST_GEOMETRY_SIGNALS;
	xGeometryRequestFresh : BOOL;
	xGeometryStopAttempt : BOOL;
	eGeometryPlace : E_POINT_NAME;
	eGeometrySafe : E_POINT_NAME;
	eGeometryChange : E_POINT_NAME;
    // Диагностика физического I/O: один владелец подмен и FIFO на 100 событий.
    axIoRawDi : ARRAY [1..84] OF BOOL;
    axIoUsedDi : ARRAY [1..84] OF BOOL;
    axIoForced : ARRAY [1..84] OF BOOL;
    axIoForceValue : ARRAY [1..84] OF BOOL;
    axIoDoForced : ARRAY [1..50] OF BOOL;
    xIoSnapshotPublishing : BOOL;
    axIoDoForceValue : ARRAY [1..50] OF BOOL;
    axIoDoInhibited : ARRAY [1..50] OF BOOL;
    axIoDoAllowed : ARRAY [1..50] OF BOOL;
    axIoDoOnAllowed : ARRAY [1..50] OF BOOL;
    axIoGripperBase : ARRAY [1..3] OF BOOL;
    axIoAutoDo : ARRAY [1..50] OF BOOL;
    axIoMagazineInvalidated : ARRAY [1..2] OF BOOL;
    xIoRawSafetyOk : BOOL;
    xIoManualActive : BOOL;
    xIoManualEndedByOperator : BOOL;
    xIoDoRejected : BOOL;
    xIoEmergencyResetRejected : BOOL;
    xIoEmergencyResetRequested : BOOL;
    udiIoEmergencyRequestSeq : UDINT;
    axIoOutput : ARRAY [1..50] OF BOOL;
    axIoPreviousRaw : ARRAY [1..84] OF BOOL;
    axIoPreviousUsed : ARRAY [1..84] OF BOOL;
    axIoPreviousOutput : ARRAY [1..50] OF BOOL;
    astIoEvent : ARRAY [1..100] OF ST_PHYSICAL_IO_EVENT;
    xIoInitialized : BOOL;
    xIoOverrideRejected : BOOL;
    xIoBusy : BOOL;
    uiIoIndex : UINT;
    uiIoWord : UINT;
    uiIoBit : UINT;
    dwIoBit : DWORD;
    udiIoNowMs : UDINT;
    udiIoLastTickMs : UDINT;
    uliIoClockMs : ULINT;
    udiIoHeartbeatSeen : UDINT;
    uliIoLeaseAgeMs : ULINT;
    tonIoOverrideWatchdog : TON;
    udiIoRequestSeq : UDINT;
    uiIoRequestAction : UINT;
    uiIoRequestIndex : UINT;
    xIoRequestValue : BOOL;
	xPhysicalNormal : BOOL;
	xPhysicalWasNormal : BOOL;
	xPhysicalInputEnable : BOOL;
	xPhysicalOutputEnable : BOOL;
	xPhysicalOutputWasEnabled : BOOL;
	uiPhysicalInput : UINT;
	tPhysicalRise : TIME;
	tPhysicalFall : TIME;
	axPhysicalRaw : ARRAY [1..84] OF BOOL;
	axPhysicalFiltered : ARRAY [1..80] OF BOOL;
	axPhysicalButtonArmed : ARRAY [1..80] OF BOOL;
	afbPhysicalInputFilter : ARRAY [1..80] OF FB_DI_FILTER;
	astMachineStatusRaw : ARRAY [1..3] OF ST_MACHINE_IO_STATUS;
	AXIS_X         : FB_AXIS; // Управление осью X
	AXIS_Y         : FB_AXIS; // Управление осью Y
	AXIS_Z         : FB_AXIS; // Управление осью Z
	GROUP_XYZ      : FB_AXIS_GROUP; // Управление группой осей XYZ
	SIMULATION_DYNAMICS : FB_SIMULATION_DYNAMIC_LIMITS; // Транзакционное масштабирование лимитов XYZ между тестами
	MOTION_MANAGER : FB_MOTION_MANAGER; // Менеджер движения по именованным точкам
	MACHINE_1      : FB_MACHINE; // Логика первого станка
	MACHINE_2      : FB_MACHINE; // Логика второго станка
	MACHINE_3      : FB_MACHINE; // Логика третьего станка
	MACHINE_1_SIM  : FB_MACHINE_SIMULATION; // Симуляция первого станка
	MACHINE_2_SIM  : FB_MACHINE_SIMULATION; // Симуляция второго станка
	MACHINE_3_SIM  : FB_MACHINE_SIMULATION; // Симуляция третьего станка
	MACHINE_1_FAULT: FB_MACHINE_FAULT_INJECTOR; // Инъекция обратной связи первого станка
	MACHINE_2_FAULT: FB_MACHINE_FAULT_INJECTOR; // Инъекция обратной связи второго станка
	MACHINE_3_FAULT: FB_MACHINE_FAULT_INJECTOR; // Инъекция обратной связи третьего станка
	TWIN_AXIS_1 : FB_AXIS;
	TWIN_AXIS_2 : FB_AXIS;
	TWIN : ARRAY [1..2] OF FB_TWO_PALLET;
	axTwinMagazineExchangeInProgress : ARRAY [1..2] OF BOOL; // Защёлка фактической смены палет для адресной блокировки магазина
	TWIN_SIM : ARRAY [1..2] OF FB_TWO_PALLET_SIMULATION;
	astTwinCommand : ARRAY [1..2] OF ST_TWO_PALLET_COMMAND;
	axTwinConfigurationChanged : ARRAY [1..2] OF BOOL;
	axTwinExternalCommandRejected : ARRAY [1..2] OF BOOL;
	audiTwinWarningSeen : ARRAY [1..2] OF UDINT;
	audiPartWarningSeen : ARRAY [1..2] OF UDINT;
	astMagazineWarningMerged : ARRAY [1..2] OF ST_WARNING_EVENT;
	uiTwin : UINT;
	uiTwinPallet : UINT;
	uiTwinRobotPalletBefore : UINT; // Смена роли после ручного восстановления снимает прежнюю готовность загрузки
	uiTwinSlot : UINT;
	udiTwinSnapshot : UDINT;
	xTwinStartup : BOOL;
	xTwinSimulationInitialized : BOOL;
	axTwinSimIoOwned : ARRAY [1..2] OF BOOL;
	axTwinSafetyBusy : ARRAY [1..2] OF BOOL;
	axButtonStationInput : ARRAY [1..4] OF BOOL; // Физическая кнопка или виртуальный вход SIMULATION
	axButtonStationEmergencyStopInput : ARRAY [1..4] OF BOOL; // Физический грибок или виртуальный вход SIMULATION
	axTwinRobotStopLatched : ARRAY [1..2] OF BOOL;
	xTwinRobotSwapWindow : BOOL;
	xTwinRobotOperation : BOOL; // Текущая, ожидающая отключения или уже выданная операция магазина
	xTwinOtherLoaded : BOOL;
	xTwinAutoSwapEnabled : BOOL;
	axTwinAutoSwapPending : ARRAY [1..2] OF BOOL; // Законченная палета ждёт окна автоматического обмена
	axMagazineInventoryChanged : ARRAY [1..2] OF BOOL; // Смена/правка только рабочего банка снимает его Finished
	xTwinInventoryCommand : BOOL;
	uiTwinRequestResult : UINT;
	stTwinRequest : ST_TWO_PALLET_REQUEST;
	fbMagazine1    : FB_MAGAZINE; // Первый статичный магазин
	fbMagazine2    : FB_MAGAZINE; // Второй статичный магазин
	ROBOT          : FB_ROBOT; // Координация движений и захвата робота
	ROBOT_MODBUS   : FB_ROBOT_MODBUS; // Modbus TCP транспорт внешнего контроллера
	TYPE_CONFIG    : FB_MULTI_TYPE_CONFIG_MANAGER; // Конфигурация типов продукции
	CELL_SAFETY    : FB_CELL_SAFETY; // Дискретный контур безопасности, двери и внешние кнопки
	CELL_MANAGER   : FB_CELL_MANAGER; // Универсальный автоматический цикл для одного-трёх типов
	ALARM_MANAGER  : FB_ALARM_MANAGER; // Журнал аварий и предупреждений
	fbAlarmHorn : FB_ALARM_HORN; // Импульс на каждую новую аварийную маску
	tonSignalTowerBlink : TON; // Полупериод мигания колонны — 500 мс
	usiSignalTowerMode : USINT; // 1 работа; 2 готова; 3 предупреждение; 4 авария; 5 не готова
	usiSignalTowerPreviousMode : USINT;
	xSignalTowerBlinkOn : BOOL := TRUE;
	uiHmiCommandIndex : UINT;
	udiHmiCommandNowMs : UDINT;
	axHmiCommandConsumed : ARRAY [1..121] OF BOOL;
	axHmiCommandWasHigh : ARRAY [1..121] OF BOOL;
	axHmiInternalPulse : ARRAY [1..121] OF BOOL; // Internal scenario events, consumed next scan
	axHmiCommandPulse : ARRAY [1..121] OF BOOL;
	audiHmiCommandSnapshot : ARRAY [1..121] OF UDINT;
	udiCellSettingSnapshot : UDINT;
	xCellSettingRejected : BOOL;
	uiMachine      : UINT; // Индекс станка при обработке команд HMI
	iDetail        : SINT; // Индекс слота при передаче состояния магазина в HMI
	xRobotHmiPermit: BOOL; // Разрешение ручных команд робота с HMI
	udiCellModeCommandSnapshot : UDINT; // Снимок маркера транзакции текущего скана
	uiCellModeRejectReason : UINT; // Одноцикловая причина отказа для журнала ячейки
	xDrivesReady   : BOOL; // Все оси и группа готовы к движению
	xDrivesPowered : BOOL; // На все три оси фактически подано питание
	xAnyDrivePowered : BOOL; // Хотя бы на одну ось фактически подано питание
	xDrivesOff     : BOOL; // Все силовые части отключены, группа в GroupDisabled
	xPowerTransitionActive : BOOL; // Выполняется последовательность включения или отключения
	xPowerDisableRequest : BOOL; // Единый запрос штатного отключения через группу
	xDriveError    : BOOL; // Активна ошибка хотя бы одной оси или группы
	xAxisDriveError : BOOL; // Активна ошибка одиночной оси; не включает административную ошибку группы
	xGroupError    : BOOL; // Активна ошибка координатной группы
	xMotionBusy    : BOOL; // Хотя бы одна ось ещё выполняет команду
	xGroupMotionBusy : BOOL; // Координатная группа выполняет движение или остановку
	xRobotAutoPowerOff : BOOL; // Автоматическое снятие питания приводов при аварии робота
	xHmiConnectionAlive : BOOL; // Watchdog связи HMI -> PLC
	xManualRecoveryActive : BOOL; // Ограниченное ручное восстановление при общей ошибке
	xHmiRobotActionBaseAllowed : BOOL; // Условия ручного перемещения робота к точке
	xHmiRobotPointTargetAllowed : BOOL; // Люк соответствующего станка открыт для входной точки
	xHmiRobotPointAllowed : BOOL; // Полное разрешение выбранной ручной точки
	eHmiRobotStatusAction : E_ROBOT_ACTION; // Действие для отображения xAllowed/reason
	eHmiRobotStatusPoint : E_POINT_NAME; // Точка для отображения xAllowed/reason
	xHmiRobotStatusPointTargetAllowed : BOOL; // Безопасность выбранной HMI-точки
	xHmiRobotStatusPointAllowed : BOOL; // Полное разрешение выбранной HMI-точки
	xHmiGripperActionBaseAllowed : BOOL; // Условия ручного действия захвата независимо от Motion-слоя
	xHmiRobotActionAllowed : BOOL;
	xHmiRobotActionAttempt : BOOL;
	rtHmiRobotAction : R_TRIG;
	udiLastHmiHeartbeat : UDINT; // Последний принятый heartbeat HMI
	tonHmiWatchdog : TON; // Таймаут HMI heartbeat
	udiLastMobileMotionHeartbeat : UDINT; // Последний heartbeat мобильной аренды
	tonMobileMotionWatchdog : TON; // Таймаут gateway/телефон -> PLC для мобильного движения
	rtMobileMotionStart : R_TRIG; // Фронт новой мобильной аренды
	xMobileMotionLeaseActive : BOOL; // PLC защёлкнул мобильного владельца до полного останова
	xMobileMotionConnectionAlive : BOOL; // Мобильный heartbeat обновляется
	xMobileMotionStopRequest : BOOL; // Независимый запрос контролируемой остановки оси
	rMobileMotionSpeedLimitPercent : REAL := 0.1; // Защёлкнутый глобальный лимит телефона
	rRobotManualEffectiveSpeedPercent : REAL := 0.1; // Итоговый override после PLC-ограничения
	uiManualAxisOwner : UINT; // Единственная ось-владелец текущей команды HMI
	uiManualAxisRequest : UINT; // Ось, запросившая новую ручную команду в текущем цикле
	axManualAxisBaseAllowed : ARRAY [1..3] OF BOOL;
	axManualAxisCommandRejected : ARRAY [1..3] OF BOOL;
	artManualAxisReject : ARRAY [1..3] OF R_TRIG;
	artHmiAxisHome : ARRAY [1..3] OF R_TRIG; // Фронты импульсных Home-команд HMI
	artHmiAxisMoveAbsolute : ARRAY [1..3] OF R_TRIG; // Фронты абсолютных команд HMI
	artHmiAxisMoveRelative : ARRAY [1..3] OF R_TRIG; // Фронты шаговых команд HMI
	axHmiAxisHomePulse : ARRAY [1..3] OF BOOL;
	axHmiAxisMoveAbsolutePulse : ARRAY [1..3] OF BOOL;
	axHmiAxisMoveRelativePulse : ARRAY [1..3] OF BOOL;
	alrRobotManualRatedVelocity : ARRAY [1..3] OF LREAL; // Фактические 100% из AXIS_REF_SM3
	alrRobotRatedAcceleration : ARRAY [1..3] OF LREAL; // Максимальное ускорение из AXIS_REF_SM3
	alrRobotRatedDeceleration : ARRAY [1..3] OF LREAL; // Максимальное замедление из AXIS_REF_SM3
	alrRobotRatedJerk : ARRAY [1..3] OF LREAL; // Максимальный jerk из AXIS_REF_SM3
	axRobotSoftwareLimitsEnabled : ARRAY [1..3] OF BOOL; // Фактическое включение software limits в AXIS_REF_SM3
	alrRobotSoftwareMinPosition : ARRAY [1..3] OF LREAL; // Отрицательный software limit SoftMotion
	alrRobotSoftwareMaxPosition : ARRAY [1..3] OF LREAL; // Положительный software limit SoftMotion
	alrRobotJogVelocity : ARRAY [1..3] OF LREAL; // Скорость одиночной оси с учётом общего коэффициента
	xHmiDrivesEnableAccepted : BOOL; // Авторитетное решение RunMotion по команде включения
	xHmiDrivesDisableAccepted : BOOL; // Авторитетное решение RunMotion по команде отключения
	xHmiResetAccepted : BOOL; // Авторитетное решение RunMotion по команде сброса
	xHmiStopAccepted : BOOL; // Авторитетное решение RunMotion по команде остановки
	xRobotMotionCommandActive : BOOL; // Принятая команда, включая проверку точки и освобождение
	xRobotProgramStopRequest : BOOL; // Штатная остановка группового движения по запросу автоматики
	xMotionResetRequest : BOOL; // Общий запрос последовательного сброса группы и осей
	xGroupResetPulse : BOOL; // Импульс MC_GroupReset; он также сбрасывает оси группы
	xAxisResetPulse : BOOL; // Последующая очистка локальных защёлок FB_AXIS
	xMotionResetBusy : BOOL; // Последовательность сброса Motion-слоя активна
	rtMotionReset : R_TRIG; // Фронт единого запроса сброса Motion-слоя
	eMotionResetState : E_MOTION_RESET_STATE := E_MOTION_RESET_STATE.IDLE;
	xAlarmResetRequired : BOOL; // Хотя бы один владелец общей команды находится в аварии
	xAlarmResetAllowed : BOOL; // Все активные владельцы аварий готовы принять общий сброс
	stRobotHmiCommand : ST_ROBOT_COMMAND; // Команда робота с учётом оперативной остановки HMI
	stSelectedMagazineCommand : ST_ROBOT_COMMAND; // Единственная команда двух магазинов роботу
	stMagazinePointCommand : ST_ROBOT_COMMAND; // Команда, по которой рассчитывается временная точка
	eMagazineBasePoint : E_POINT_NAME; // База выбранного магазина
	uiMagazine : UINT; // Индекс магазина 1..2
	auiMagazineEditSlot : ARRAY [1..2] OF UINT; // Новый контракт с fallback на legacy-команду первого магазина
	astMachineFaultRequest : ARRAY [1..3] OF ST_MACHINE_FAULT_REQUEST; // Запросы ошибок станков
	astAxisFaultRequest    : ARRAY [1..3] OF ST_AXIS_FAULT_REQUEST; // Запросы ошибок осей
	stAxisGroupFaultRequest: ST_AXIS_GROUP_FAULT_REQUEST; // Запрос ошибки группы XYZ
	stRobotFaultRequest    : ST_ROBOT_FAULT_REQUEST; // Запросы ошибок робота и точки
	astMagazineFaultRequest : ARRAY [1..2] OF ST_MAGAZINE_FAULT_REQUEST; // Диагностика двух магазинов
	stCellFaultRequest     : ST_CELL_FAULT_REQUEST; // Запрос локальной ошибки менеджера ячейки
	stSafetyFaultRequest   : ST_CELL_SAFETY_FAULT_REQUEST; // Независимые инъекции дискретной безопасности
	astAlarmSource : ARRAY [1..19] OF ST_ALARM_SOURCE_DATA; // Старые коды сохранены; ГК 1/2 добавлены в конец
	astAdditionalCellWarning : ARRAY [1..2] OF ST_WARNING_EVENT; // 1: конфигуратор, 2: общие предупреждения ГК
	uiPointEditorIndex : UINT; // Компактный индекс фиксированной точки редактора 1..14
	uiPointEditorGeometryStation : UINT; // 0 прежняя точка, 1/2 база ГК
	uiPointStorageIndex : UINT; // Индекс в совместимом Persistent-массиве 1..15
	ePointEditorName : E_POINT_NAME; // Фактический enum выбранной инженерной точки
	xPointTableReady : BOOL; // Все 12 базовых точек подтверждены редактором
	axMachinePointsReady : ARRAY [1..3] OF BOOL; // Три рабочие точки каждого станка
	axMagazinePointsReady : ARRAY [1..2] OF BOOL; // База и оба Z-смещения каждого магазина
	xCellPointsReady : BOOL; // HOME_SAFETY и точки только включённого оборудования
	xPointEditorBaseAllowed : BOOL; // Общие безопасные условия Capture/Save
	xPointEditorAllHomed : BOOL; // Все оси XYZ прошли Home
	xPointEditorRequestValid : BOOL; // Индекс и код новой транзакции распознаны
	xPointEditorDraftValid : BOOL; // XYZ и скорость черновика прошли проверку
	xPointEditorMagazinePoint : BOOL; // Выбрана базовая точка магазина 1 или 2
	xPointEditorGeometrySave : BOOL; // SAVE базы ГК не зависит от технологических блокировок
	udiLastPointEditorCommandSeq : UDINT; // Последняя обработанная транзакция редактора
	xPointCheckRequest : BOOL;
	xPointCheckActive : BOOL;
	xPointCheckStopping : BOOL;
	xPointCheckSeenBusy : BOOL;
	xPointCheckSeenDone : BOOL; // Терминальный ответ Motion хранится до фактического останова
	xPointCheckStopRequest : BOOL;
	xPointCheckConnectionAlive : BOOL;
	udiLastPointCheckHeartbeat : UDINT;
	tonPointCheckWatchdog : TON;
	tonPointCheckStart : TON;
	ePointCheckName : E_POINT_NAME;
	uiPointCheckLoop : UINT;
	uiPointCheckMachine : UINT;
	uiPointCheckReason : UINT;
	stPointCheckCandidate : ST_POINT;
	rPointCheckLatchedSpeed : REAL;
	lrGroupVelocityOverride : LREAL;
	xRobotInterfaceReady : BOOL; // Готовность применённого интерфейса робота
	lrRobotActualX : LREAL; // Координаты выбранного источника управления
	lrRobotActualY : LREAL;
	lrRobotActualZ : LREAL;
	xModeCommonSafe : BOOL; // Общие условия изменения источника управления
	xAllMachinesIdle : BOOL;
	rtRobotModeApply : R_TRIG;
	rtModbusSettingsApply : R_TRIG;
	xModbusHmiInitialized : BOOL;
	uiRobotInterfaceWarningCode : UINT;
	uiRobotManualMagazineIndex : UINT;
	uiRobotManualMagazineRow : UINT;
	uiRobotManualMagazineColumn : UINT;
	rtTestEnvironmentApply : R_TRIG;
	rtTestSpeedProfileApply : R_TRIG;
	rtTestScenarioApply : R_TRIG;
	xTestInitializePulse : BOOL;
	xTestAbortActive : BOOL; // Тестовая отмена действует только в виртуальной среде
	xTestStable : BOOL;
	xTestScenarioValid : BOOL;
	uiTestIndex : UINT;
	uiTestMagazine : UINT;
	uiTestFaultOwnerCount : UINT;
	adwTestMagazineFaultMask : ARRAY [1..2] OF DWORD;
	xApplicationStartupInitialized : BOOL; // Однократная инициализация безопасных настроек после старта/Online Change
END_VAR

VAR CONSTANT
	WRN_HMI_MANUAL_REJECTED : UINT := 12; // PLC отклонил команду расширенного ручного управления
	WRN_ROBOT_MODE_REJECTED : UINT := 13; // PLC отклонил переключение источника управления
	WRN_MODBUS_SETTINGS_REJECTED : UINT := 14; // PLC отклонил применение параметров соединения
	WRN_POINT_EDIT_REJECTED : UINT := 15; // PLC отклонил Capture/Save инженерной точки
	WRN_POINT_CHECK_REJECTED : UINT := 16; // Проверка точки отклонена
	WRN_POINT_CHECK_INTERRUPTED : UINT := 17; // Проверка остановлена потерей связи/разрешений
	aePointCheckNames : ARRAY [1..14] OF E_POINT_NAME := [
		E_POINT_NAME.MACHINE_1_ABOVE, E_POINT_NAME.MACHINE_1_CHUCK_APROACH, E_POINT_NAME.MACHINE_1_CHUCK_POSITION,
		E_POINT_NAME.MACHINE_2_ABOVE, E_POINT_NAME.MACHINE_2_CHUCK_APROACH, E_POINT_NAME.MACHINE_2_CHUCK_POSITION,
		E_POINT_NAME.MACHINE_3_ABOVE, E_POINT_NAME.MACHINE_3_CHUCK_APROACH, E_POINT_NAME.MACHINE_3_CHUCK_POSITION,
		E_POINT_NAME.HOME_SAFETY, E_POINT_NAME.MAGAZINE_1_DETAIL, E_POINT_NAME.MAGAZINE_2_DETAIL,
		E_POINT_NAME.GEOMETRY_1_PLACE, E_POINT_NAME.GEOMETRY_2_PLACE];
	alrRobotManualFallbackVelocity : ARRAY [1..3] OF LREAL := [1000.0, 1000.0, 1000.0]; // Резерв, если привод не публикует динамический предел
	alrRobotManualAcceleration : ARRAY [1..3] OF LREAL := [1000.0, 1000.0, 1000.0]; // Резерв ускорения, если привод не публикует предел
	alrRobotManualDeceleration : ARRAY [1..3] OF LREAL := [1000.0, 1000.0, 1000.0]; // Резерв замедления, если привод не публикует предел
	alrRobotManualJerk : ARRAY [1..3] OF LREAL := [10000.0, 10000.0, 10000.0]; // Резерв jerk, если привод не публикует предел
END_VAR

SetApplicationDefaults();
ReadHmiCommands();
ReadHmiInputs();
ReadIoEmergencyStop();
ReadPhysicalInputs();
RunSafety();
ResetIoEmergencyStop();
RunMotion();
RunRobotModbus();
RunTestControl();
RunTwoPallet();
RunGeometryControl();
RunCellControl();
RunMachines();
RunMagazine();
RunTwoPalletAxis();
RunRobot();
RunAlarms();
RunSignalTower();
WritePhysicalOutputs();
RecordIoDiagnostics();
PublishGeometryControl();
PublishHmi();

METHOD PRIVATE ReadHmiInputs
// HMI обязана поддерживать heartbeat. При потере связи PLC снимает только
// расширенные ручные команды; технологические проверки ниже остаются в PLC.
tonHmiWatchdog(
	IN := GVL_HMI.udiHmiHeartbeat = udiLastHmiHeartbeat,
	PT := GVL_CELL_SETTINGS.tHmiWatchdogTimeout
);
IF GVL_HMI.udiHmiHeartbeat <> udiLastHmiHeartbeat THEN
	udiLastHmiHeartbeat := GVL_HMI.udiHmiHeartbeat;
END_IF;
xHmiConnectionAlive := NOT tonHmiWatchdog.Q;

// Мобильная аренда отделена от общего HMI heartbeat. Gateway может быть жив,
// но движение обязано остановиться, если телефон перестал подтверждать аренду.
rtMobileMotionStart(CLK := GVL_HMI.xMobileMotionActive);
tonMobileMotionWatchdog(
	IN := GVL_HMI.xMobileMotionActive
		AND (GVL_HMI.udiMobileMotionHeartbeat = udiLastMobileMotionHeartbeat),
	PT := GVL_CELL_SETTINGS.tMobileMotionWatchdogTimeout
);
IF GVL_HMI.udiMobileMotionHeartbeat <> udiLastMobileMotionHeartbeat THEN
	udiLastMobileMotionHeartbeat := GVL_HMI.udiMobileMotionHeartbeat;
END_IF;
IF rtMobileMotionStart.Q THEN
	xMobileMotionLeaseActive := TRUE;
	rMobileMotionSpeedLimitPercent := LIMIT(
		REAL#0.1,
		GVL_CELL_SETTINGS.rPointCheckSpeedPercent,
		REAL#100.0
	);
END_IF;
IF xMobileMotionLeaseActive THEN
	// Во время аренды лимит разрешено только уменьшать. Повышение настройки
	// применяется уже к следующему мобильному движению.
	rMobileMotionSpeedLimitPercent := MIN(
		rMobileMotionSpeedLimitPercent,
		LIMIT(REAL#0.1, GVL_CELL_SETTINGS.rPointCheckSpeedPercent, REAL#100.0)
	);
END_IF;
xMobileMotionConnectionAlive := GVL_HMI.xMobileMotionActive
	AND NOT tonMobileMotionWatchdog.Q;
xMobileMotionStopRequest := xMobileMotionLeaseActive
	AND (NOT GVL_HMI.xMobileMotionActive
		OR NOT xMobileMotionConnectionAlive
		OR NOT xHmiConnectionAlive);
IF xMobileMotionStopRequest THEN
	// Сбрасываем вход аренды в PLC: восстановление сети не может само возобновить ход.
	GVL_HMI.xMobileMotionActive := FALSE;
	FOR uiMachine := 1 TO 3 DO
		GVL_HMI.astAxisHmiCommand[uiMachine].xJogPositive := FALSE;
		GVL_HMI.astAxisHmiCommand[uiMachine].xJogNegative := FALSE;
	END_FOR;
END_IF;
GVL_HMI.xMobileMotionLeaseAlive := xMobileMotionLeaseActive
	AND xMobileMotionConnectionAlive
	AND NOT xMobileMotionStopRequest;
GVL_HMI.rMobileMotionAppliedSpeedPercent := rMobileMotionSpeedLimitPercent;

xPointCheckRequest := FALSE;
tonPointCheckWatchdog(
	IN := GVL_HMI.udiPointCheckHeartbeat = udiLastPointCheckHeartbeat,
	PT := GVL_CELL_SETTINGS.tPointCheckWatchdogTimeout
);
IF GVL_HMI.udiPointCheckHeartbeat <> udiLastPointCheckHeartbeat THEN
	udiLastPointCheckHeartbeat := GVL_HMI.udiPointCheckHeartbeat;
END_IF;
xPointCheckConnectionAlive := (udiLastPointCheckHeartbeat <> UDINT#0) AND NOT tonPointCheckWatchdog.Q;
xPointCheckStopRequest := xPointCheckActive AND (GVL_HMI.xPointCheckStop
	OR NOT xPointCheckConnectionAlive OR NOT xHmiConnectionAlive);
// Stop is a PLC-owned one-scan event; its request counter is never cleared here.

